  MoveL 1290 to (-200, -11.4, 56.6) mm, rotated rx 180 ry 0 rz 180 deg; joints [-15.315, -59.69, 128.134, 163.594, 69.246, -84.044]
  MoveL 1291 to (-200, -12, 56.6) mm, rotated rx 180 ry 0 rz 180 deg; joints [-15.315, -59.729, 128.133, 163.589, 69.207, -84.031]
  MoveL 1292 to (0, -12, 56.6) mm, rotated rx 180 ry 0 rz 180 deg; joints [-13.166, -51.617, 112.007, 164.94, 61.242, -82.624]
  MoveL 1293 to (0, -12.6, 56.6) mm, rotated rx 180 ry 0 rz 180 deg; joints [-13.166, -51.649, 112.006, 164.936, 61.21, -82.614]
  MoveL 1294 to (-200, -12.6, 56.6) mm, rotated rx 180 ry 0 rz 180 deg; joints [-15.315, -59.768, 128.131, 163.585, 69.169, -84.019]
  MoveL 1295 to (-200, -13.2, 56.6) mm, rotated rx 180 ry 0 rz 180 deg; joints [-15.315, -59.807, 128.13, 163.581, 69.13, -84.007]
  MoveL 1296 to (0, -13.2, 56.6) mm, rotated rx 180 ry 0 rz 180 deg; joints [-13.166, -51.681, 112.005, 164.931, 61.178, -82.605]
  MoveL 1297 to (0, -13.8, 56.6) mm, rotated rx 180 ry 0 rz 180 deg; joints [-13.166, -51.713, 112.003, 164.926, 61.146, -82.595]
  MoveL 1298 to (-200, -13.8, 56.6) mm, rotated rx 180 ry 0 rz 180 deg; joints [-15.315, -59.846, 128.129, 163.576, 69.091, -83.995]
  MoveL 1299 to (-200, -14.4, 56.6) mm, rotated rx 180 ry 0 rz 180 deg; joints [-15.315, -59.885, 128.127, 163.572, 69.052, -83.982]
  MoveL 1300 to (0, -14.4, 56.6) mm, rotated rx 180 ry 0 rz 180 deg; joints [-13.166, -51.745, 112.002, 164.921, 61.114, -82.585]
  MoveL 1301 to (0, -15, 56.6) mm, rotated rx 180 ry 0 rz 180 deg; joints [-13.166, -51.776, 112.001, 164.917, 61.082, -82.575]
  MoveL 1302 to (-200, -15, 56.6) mm, rotated rx 180 ry 0 rz 180 deg; joints [-15.315, -59.924, 128.126, 163.567, 69.013, -83.97]
  MoveL 1303 to (-200, -15.6, 56.6) mm, rotated rx 180 ry 0 rz 180 deg; joints [-15.315, -59.963, 128.124, 163.563, 68.975, -83.958]
  MoveL 1304 to (0, -15.6, 56.6) mm, rotated rx 180 ry 0 rz 180 deg; joints [-13.166, -51.808, 111.999, 164.912, 61.05, -82.565]
  MoveL 1305 to (0, -16.2, 56.6) mm, rotated rx 180 ry 0 rz 180 deg; joints [-13.166, -51.84, 111.998, 164.907, 61.018, -82.555]
  MoveL 1306 to (-200, -16.2, 56.6) mm, rotated rx 180 ry 0 rz 180 deg; joints [-15.315, -60.001, 128.122, 163.559, 68.936, -83.946]
  MoveL 1307 to (-200, -16.8, 56.6) mm, rotated rx 180 ry 0 rz 180 deg; joints [-15.315, -60.04, 128.121, 163.554, 68.897, -83.933]
  MoveL 1308 to (0, -16.8, 56.6) mm, rotated rx 180 ry 0 rz 180 deg; joints [-13.166, -51.872, 111.996, 164.902, 60.986, -82.545]
  MoveL 1309 to (0, -17.4, 56.6) mm, rotated rx 180 ry 0 rz 180 deg; joints [-13.166, -51.903, 111.995, 164.898, 60.954, -82.535]
  MoveL 1310 to (-200, -17.4, 56.6) mm, rotated rx 180 ry 0 rz 180 deg; joints [-15.315, -60.079, 128.119, 163.55, 68.858, -83.921]
  MoveL 1311 to (-200, -18, 56.6) mm, rotated rx 180 ry 0 rz 180 deg; joints [-15.315, -60.118, 128.117, 163.545, 68.819, -83.909]
  MoveL 1312 to (0, -18, 56.6) mm, rotated rx 180 ry 0 rz 180 deg; joints [-13.166, -51.935, 111.993, 164.893, 60.922, -82.526]
  MoveL 1313 to (0, -18.6, 56.6) mm, rotated rx 180 ry 0 rz 180 deg; joints [-13.166, -51.967, 111.992, 164.888, 60.89, -82.516]
  MoveL 1314 to (-200, -18.6, 56.6) mm, rotated rx 180 ry 0 rz 180 deg; joints [-15.315, -60.157, 128.116, 163.541, 68.78, -83.896]
  MoveL 1315 to (-200, -19.2, 56.6) mm, rotated rx 180 ry 0 rz 180 deg; joints [-15.315, -60.196, 128.114, 163.536, 68.741, -83.884]
  MoveL 1316 to (0, -19.2, 56.6) mm, rotated rx 180 ry 0 rz 180 deg; joints [-13.166, -51.998, 111.99, 164.883, 60.858, -82.506]
  MoveL 1317 to (0, -19.8, 56.6) mm, rotated rx 180 ry 0 rz 180 deg; joints [-13.166, -52.03, 111.988, 164.878, 60.826, -82.496]
  MoveL 1318 to (-200, -19.8, 56.6) mm, rotated rx 180 ry 0 rz 180 deg; joints [-15.315, -60.235, 128.112, 163.532, 68.702, -83.872]
  MoveL 1319 to (-200, -20.4, 56.6) mm, rotated rx 180 ry 0 rz 180 deg; joints [-15.315, -60.273, 128.11, 163.527, 68.663, -83.859]
  MoveL 1320 to (0, -20.4, 56.6) mm, rotated rx 180 ry 0 rz 180 deg; joints [-13.166, -52.062, 111.987, 164.873, 60.794, -82.486]
  MoveL 1321 to (0, -21, 56.6) mm, rotated rx 180 ry 0 rz 180 deg; joints [-13.166, -52.093, 111.985, 164.869, 60.762, -82.476]
  MoveL 1322 to (-200, -21, 56.6) mm, rotated rx 180 ry 0 rz 180 deg; joints [-15.315, -60.312, 128.108, 163.523, 68.624, -83.847]
  MoveL 1323 to (-200, -21.6, 56.6) mm, rotated rx 180 ry 0 rz 180 deg; joints [-15.315, -60.351, 128.107, 163.518, 68.585, -83.835]
  MoveL 1324 to (0, -21.6, 56.6) mm, rotated rx 180 ry 0 rz 180 deg; joints [-13.166, -52.125, 111.983, 164.864, 60.729, -82.466]
  MoveL 1325 to (0, -22.2, 56.6) mm, rotated rx 180 ry 0 rz 180 deg; joints [-13.166, -52.156, 111.982, 164.859, 60.697, -82.456]
  MoveL 1326 to (-200, -22.2, 56.6) mm, rotated rx 180 ry 0 rz 180 deg; joints [-15.315, -60.39, 128.105, 163.514, 68.546, -83.822]
  MoveL 1327 to (-200, -22.8, 56.6) mm, rotated rx 180 ry 0 rz 180 deg; joints [-15.315, -60.428, 128.103, 163.509, 68.507, -83.81]
  MoveL 1328 to (0, -22.8, 56.6) mm, rotated rx 180 ry 0 rz 180 deg; joints [-13.166, -52.188, 111.98, 164.854, 60.665, -82.446]
  MoveL 1329 to (0, -23.4, 56.6) mm, rotated rx 180 ry 0 rz 180 deg; joints [-13.166, -52.219, 111.978, 164.849, 60.633, -82.436]
  MoveL 1330 to (-200, -23.4, 56.6) mm, rotated rx 180 ry 0 rz 180 deg; joints [-15.315, -60.467, 128.101, 163.505, 68.468, -83.797]
  MoveL 1331 to (-200, -24, 56.6) mm, rotated rx 180 ry 0 rz 180 deg; joints [-15.315, -60.506, 128.099, 163.5, 68.429, -83.785]
  MoveL 1332 to (0, -24, 56.6) mm, rotated rx 180 ry 0 rz 180 deg; joints [-13.166, -52.251, 111.976, 164.844, 60.601, -82.426]
  MoveL 1333 to (0, -24.6, 56.6) mm, rotated rx 180 ry 0 rz 180 deg; joints [-13.166, -52.282, 111.974, 164.839, 60.568, -82.416]
  MoveL 1334 to (-200, -24.6, 56.6) mm, rotated rx 180 ry 0 rz 180 deg; joints [-15.315, -60.545, 128.097, 163.496, 68.39, -83.772]
  MoveL 1335 to (-200, -25.2, 56.6) mm, rotated rx 180 ry 0 rz 180 deg; joints [-15.315, -60.583, 128.095, 163.491, 68.351, -83.76]
  MoveL 1336 to (0, -25.2, 56.6) mm, rotated rx 180 ry 0 rz 180 deg; joints [-13.166, -52.314, 111.973, 164.834, 60.536, -82.406]
  MoveL 1337 to (0, -25.8, 56.6) mm, rotated rx 180 ry 0 rz 180 deg; joints [-13.166, -52.345, 111.971, 164.829, 60.504, -82.396]
  MoveL 1338 to (-200, -25.8, 56.6) mm, rotated rx 180 ry 0 rz 180 deg; joints [-15.315, -60.622, 128.092, 163.486, 68.312, -83.748]
  MoveL 1339 to (-200, -26.4, 56.6) mm, rotated rx 180 ry 0 rz 180 deg; joints [-15.315, -60.66, 128.09, 163.482, 68.273, -83.735]
  MoveL 1340 to (0, -26.4, 56.6) mm, rotated rx 180 ry 0 rz 180 deg; joints [-13.166, -52.377, 111.969, 164.824, 60.472, -82.386]
  MoveL 1341 to (0, -27, 56.6) mm, rotated rx 180 ry 0 rz 180 deg; joints [-13.166, -52.408, 111.967, 164.819, 60.439, -82.376]
  MoveL 1342 to (-200, -27, 56.6) mm, rotated rx 180 ry 0 rz 180 deg; joints [-15.315, -60.699, 128.088, 163.477, 68.234, -83.723]
  MoveL 1343 to (-200, -27.6, 56.6) mm, rotated rx 180 ry 0 rz 180 deg; joints [-15.315, -60.738, 128.086, 163.472, 68.195, -83.71]
  MoveL 1344 to (0, -27.6, 56.6) mm, rotated rx 180 ry 0 rz 180 deg; joints [-13.166, -52.44, 111.965, 164.814, 60.407, -82.366]
  MoveL 1345 to (0, -28.2, 56.6) mm, rotated rx 180 ry 0 rz 180 deg; joints [-13.166, -52.471, 111.963, 164.809, 60.375, -82.356]
  MoveL 1346 to (-200, -28.2, 56.6) mm, rotated rx 180 ry 0 rz 180 deg; joints [-15.315, -60.776, 128.084, 163.468, 68.156, -83.698]
  MoveL 1347 to (-200, -28.8, 56.6) mm, rotated rx 180 ry 0 rz 180 deg; joints [-15.315, -60.815, 128.081, 163.463, 68.116, -83.685]
  MoveL 1348 to (0, -28.8, 56.6) mm, rotated rx 180 ry 0 rz 180 deg; joints [-13.166, -52.503, 111.961, 164.804, 60.343, -82.346]
  MoveL 1349 to (0, -29.4, 56.6) mm, rotated rx 180 ry 0 rz 180 deg; joints [-13.166, -52.534, 111.959, 164.799, 60.31, -82.335]
  MoveL 1350 to (-200, -29.4, 56.6) mm, rotated rx 180 ry 0 rz 180 deg; joints [-15.315, -60.853, 128.079, 163.458, 68.077, -83.672]
  MoveL 1351 to (-200, -30, 56.6) mm, rotated rx 180 ry 0 rz 180 deg; joints [-15.315, -60.892, 128.077, 163.454, 68.038, -83.66]
  MoveL 1352 to (0, -30, 56.6) mm, rotated rx 180 ry 0 rz 180 deg; joints [-13.166, -52.565, 111.956, 164.794, 60.278, -82.325]
  MoveL 1353 to (0, -30.6, 56.58) mm, rotated rx 177.04 ry 0 rz 180 deg; joints [-13.235, -53.54, 111.838, 164.547, 59.233, -84.915]
  MoveL 1354 to (-200, -30.6, 56.58) mm, rotated rx 177.04 ry 0 rz 180 deg; joints [-15.394, -62.091, 127.948, 163.21, 66.774, -86.179]
  MoveL 1355 to (-200, -31.2, 56.54) mm, rotated rx 174.07 ry 0 rz 180 deg; joints [-15.428, -63.285, 127.806, 163.002, 65.501, -88.702]
  MoveL 1356 to (0, -31.2, 56.54) mm, rotated rx 174.07 ry 0 rz 180 deg; joints [-13.265, -54.511, 111.709, 164.333, 58.178, -87.515]
  MoveL 1357 to (0, -31.79, 56.46) mm, rotated rx 171.11 ry 0 rz 180 deg; joints [-13.255, -55.475, 111.57, 164.155, 57.114, -90.13]
  MoveL 1358 to (-200, -31.79, 56.46) mm, rotated rx 171.11 ry 0 rz 180 deg; joints [-15.417, -64.469, 127.651, 162.829, 64.219, -91.237]
  MoveL 1359 to (-200, -32.38, 56.35) mm, rotated rx 168.15 ry 0 rz 180 deg; joints [-15.36, -65.641, 127.484, 162.694, 62.932, -93.784]
  MoveL 1360 to (0, -32.38, 56.35) mm, rotated rx 168.15 ry 0 rz 180 deg; joints [-13.206, -56.43, 111.42, 164.013, 56.044, -92.762]
  MoveL 1361 to (0, -32.97, 56.21) mm, rotated rx 165.18 ry 0 rz 180 deg; joints [-13.118, -57.374, 111.26, 163.909, 54.969, -95.416]
  MoveL 1362 to (-200, -32.97, 56.21) mm, rotated rx 165.18 ry 0 rz 180 deg; joints [-15.259, -66.799, 127.305, 162.598, 61.643, -96.351]
  MoveL 1363 to (-200, -33.54, 56.05) mm, rotated rx 162.22 ry 0 rz 180 deg; joints [-15.112, -67.937, 127.115, 162.543, 60.354, -98.94]
  MoveL 1364 to (0, -33.54, 56.05) mm, rotated rx 162.22 ry 0 rz 180 deg; joints [-12.99, -58.304, 111.092, 163.846, 53.893, -98.094]
  MoveL 1365 to (0, -34.11, 55.85) mm, rotated rx 159.25 ry 0 rz 180 deg; joints [-12.824, -59.217, 110.914, 163.824, 52.818, -100.802]
  MoveL 1366 to (-200, -34.11, 55.85) mm, rotated rx 159.25 ry 0 rz 180 deg; joints [-14.921, -69.055, 126.916, 162.531, 59.067, -101.556]
  MoveL 1367 to (-200, -34.66, 55.62) mm, rotated rx 156.29 ry 0 rz 180 deg; joints [-14.686, -70.148, 126.706, 162.564, 57.786, -104.204]
  MoveL 1368 to (0, -34.66, 55.62) mm, rotated rx 156.29 ry 0 rz 180 deg; joints [-12.619, -60.112, 110.729, 163.847, 51.745, -103.542]
  MoveL 1369 to (0, -35.21, 55.37) mm, rotated rx 153.33 ry 0 rz 180 deg; joints [-12.376, -60.986, 110.538, 163.916, 50.677, -106.317]
  MoveL 1370 to (-200, -35.21, 55.37) mm, rotated rx 153.33 ry 0 rz 180 deg; joints [-14.406, -71.215, 126.489, 162.644, 56.513, -106.888]
  MoveL 1371 to (-200, -35.74, 55.08) mm, rotated rx 150.36 ry 0 rz 180 deg; joints [-14.083, -72.253, 126.264, 162.774, 55.251, -109.614]
  MoveL 1372 to (0, -35.74, 55.08) mm, rotated rx 150.36 ry 0 rz 180 deg; joints [-12.095, -61.837, 110.34, 164.034, 49.618, -109.135]
  MoveL 1373 to (0, -36.25, 54.77) mm, rotated rx 147.4 ry 0 rz 180 deg; joints [-11.777, -62.663, 110.136, 164.203, 48.57, -111.996]
  MoveL 1374 to (-200, -36.25, 54.77) mm, rotated rx 147.4 ry 0 rz 180 deg; joints [-13.716, -73.26, 126.033, 162.958, 54.004, -112.386]
  MoveL 1375 to (-200, -36.75, 54.44) mm, rotated rx 144.44 ry 0 rz 180 deg; joints [-13.307, -74.233, 125.797, 163.198, 52.775, -115.211]
  MoveL 1376 to (0, -36.75, 54.44) mm, rotated rx 144.44 ry 0 rz 180 deg; joints [-11.422, -63.463, 109.929, 164.427, 47.535, -114.907]
  MoveL 1377 to (0, -37.23, 54.08) mm, rotated rx 141.47 ry 0 rz 180 deg; joints [-11.032, -64.234, 109.719, 164.709, 46.517, -117.871]
  MoveL 1378 to (-200, -37.23, 54.08) mm, rotated rx 141.47 ry 0 rz 180 deg; joints [-12.856, -75.17, 125.557, 163.498, 51.566, -118.091]
  MoveL 1379 to (-200, -37.69, 53.69) mm, rotated rx 138.51 ry 0 rz 180 deg; joints [-12.364, -76.07, 125.315, 163.86, 50.381, -121.035]
  MoveL 1380 to (0, -37.69, 53.69) mm, rotated rx 138.51 ry 0 rz 180 deg; joints [-10.606, -64.975, 109.506, 165.05, 45.518, -120.893]
  MoveL 1381 to (0, -38.12, 53.28) mm, rotated rx 135.55 ry 0 rz 180 deg; joints [-10.146, -65.683, 109.292, 165.455, 44.542, -123.977]
  MoveL 1382 to (-200, -38.12, 53.28) mm, rotated rx 135.55 ry 0 rz 180 deg; joints [-11.832, -76.929, 125.071, 164.29, 49.223, -124.044]
  MoveL 1383 to (-200, -38.54, 52.85) mm, rotated rx 132.58 ry 0 rz 180 deg; joints [-11.261, -77.748, 124.828, 164.789, 48.098, -127.125]
  MoveL 1384 to (0, -38.54, 52.85) mm, rotated rx 132.58 ry 0 rz 180 deg; joints [-9.653, -66.359, 109.079, 165.925, 43.592, -127.125]
  MoveL 1385 to (0, -38.94, 52.4) mm, rotated rx 129.62 ry 0 rz 180 deg; joints [-9.128, -66.999, 108.867, 166.464, 42.671, -130.343]
  MoveL 1386 to (-200, -38.94, 52.4) mm, rotated rx 129.62 ry 0 rz 180 deg; joints [-10.652, -78.523, 124.586, 165.362, 47.007, -130.282]
  MoveL 1387 to (-200, -39.31, 51.92) mm, rotated rx 126.66 ry 0 rz 180 deg; joints [-10.007, -79.254, 124.348, 166.011, 45.956, -133.518]
  MoveL 1388 to (0, -39.31, 51.92) mm, rotated rx 126.66 ry 0 rz 180 deg; joints [-8.572, -67.603, 108.657, 167.074, 41.783, -133.633]
  MoveL 1389 to (0, -39.65, 51.44) mm, rotated rx 123.69 ry 0 rz 180 deg; joints [-7.986, -68.17, 108.45, 167.758, 40.932, -136.998]
  MoveL 1390 to (-200, -39.65, 51.44) mm, rotated rx 123.69 ry 0 rz 180 deg; joints [-9.326, -79.939, 124.113, 166.739, 44.949, -136.839]
  MoveL 1391 to (-200, -39.97, 50.93) mm, rotated rx 120.73 ry 0 rz 180 deg; joints [-8.612, -80.576, 123.885, 167.549, 43.99, -140.244]
  MoveL 1392 to (0, -39.97, 50.93) mm, rotated rx 120.73 ry 0 rz 180 deg; joints [-7.372, -68.697, 108.249, 168.515, 40.122, -140.44]
  MoveL 1393 to (0, -40.26, 50.4) mm, rotated rx 117.77 ry 0 rz 180 deg; joints [-6.731, -69.186, 108.053, 169.348, 39.355, -143.96]
  MoveL 1394 to (-200, -40.26, 50.4) mm, rotated rx 117.77 ry 0 rz 180 deg; joints [-7.867, -81.165, 123.663, 168.441, 43.084, -143.739]
  MoveL 1395 to (-200, -40.53, 49.87) mm, rotated rx 114.8 ry 0 rz 180 deg; joints [-7.091, -81.704, 123.45, 169.417, 42.234, -147.323]
  MoveL 1396 to (0, -40.53, 49.87) mm, rotated rx 114.8 ry 0 rz 180 deg; joints [-6.066, -69.633, 107.864, 170.256, 38.636, -147.559]
  MoveL 1397 to (0, -40.77, 49.31) mm, rotated rx 111.84 ry 0 rz 180 deg; joints [-5.378, -70.039, 107.683, 171.238, 37.97, -151.235]
  MoveL 1398 to (-200, -40.77, 49.31) mm, rotated rx 111.84 ry 0 rz 180 deg; joints [-6.288, -82.193, 123.246, 170.475, 41.447, -150.994]
  MoveL 1399 to (-200, -40.98, 48.75) mm, rotated rx 108.87 ry 0 rz 180 deg; joints [-5.46, -82.631, 123.053, 171.615, 40.726, -154.752]
  MoveL 1400 to (0, -40.98, 48.75) mm, rotated rx 108.87 ry 0 rz 180 deg; joints [-4.668, -70.402, 107.511, 172.293, 37.359, -154.987]
  MoveL 1401 to (0, -41.16, 48.18) mm, rotated rx 105.91 ry 0 rz 180 deg; joints [-3.939, -70.723, 107.349, 173.417, 36.808, -158.81]
  MoveL 1402 to (-200, -41.16, 48.18) mm, rotated rx 105.91 ry 0 rz 180 deg; joints [-4.608, -83.016, 122.871, 172.831, 40.077, -158.592]
  MoveL 1403 to (-200, -41.3, 47.6) mm, rotated rx 102.95 ry 0 rz 180 deg; joints [-3.736, -83.349, 122.703, 174.121, 39.502, -162.51]
  MoveL 1404 to (0, -41.3, 47.6) mm, rotated rx 102.95 ry 0 rz 180 deg; joints [-3.192, -71, 107.198, 174.605, 36.319, -162.701]
  MoveL 1405 to (0, -41.42, 47.01) mm, rotated rx 99.98 ry 0 rz 180 deg; joints [-2.431, -71.233, 107.058, 175.851, 35.897, -166.654]
  MoveL 1406 to (-200, -41.42, 47.01) mm, rotated rx 99.98 ry 0 rz 180 deg; joints [-2.845, -83.628, 122.548, 175.477, 39.007, -166.499]
  MoveL 1407 to (-200, -41.51, 46.42) mm, rotated rx 97.02 ry 0 rz 180 deg; joints [-1.94, -83.854, 122.408, 176.889, 38.595, -170.548]
  MoveL 1408 to (0, -41.51, 46.42) mm, rotated rx 97.02 ry 0 rz 180 deg; joints [-1.657, -71.421, 106.931, 177.148, 35.543, -170.659]
  MoveL 1409 to (0, -41.57, 45.82) mm, rotated rx 94.06 ry 0 rz 180 deg; joints [-0.873, -71.565, 106.816, 178.488, 35.261, -174.71]
  MoveL 1410 to (-200, -41.57, 45.82) mm, rotated rx 94.06 ry 0 rz 180 deg; joints [-1.022, -84.026, 122.283, 178.35, 38.268, -174.649]
  MoveL 1411 to (-200, -41.6, 45.22) mm, rotated rx 91.09 ry 0 rz 180 deg; joints [-0.094, -84.144, 122.173, 179.847, 38.029, -178.787]
  MoveL 1412 to (0, -41.6, 45.22) mm, rotated rx 91.09 ry 0 rz 180 deg; joints [-0.08, -71.664, 106.715, 179.86, 35.052, -178.793]
  MoveL 1413 to (0, -41.6, 44.62) mm, rotated rx 90 ry 0 rz 180 deg; joints [0.229, -71.689, 106.681, -179.6, 34.993, 179.672]
  MoveL 1414 to (-200, -41.6, 44.62) mm, rotated rx 90 ry 0 rz 180 deg; joints [0.268, -84.174, 122.137, -179.564, 37.964, 179.656]
  MoveL 1415 to (-200, -41.6, 44.02) mm, rotated rx 90 ry 0 rz 180 deg; joints [0.298, -84.174, 122.137, -179.516, 37.964, 179.618]
  MoveL 1416 to (0, -41.6, 44.02) mm, rotated rx 90 ry 0 rz 180 deg; joints [0.254, -71.689, 106.681, -179.556, 34.993, 179.637]
  MoveL 1417 to (0, -41.6, 43.42) mm, rotated rx 90 ry 0 rz 180 deg; joints [0.279, -71.688, 106.681, -179.513, 34.994, 179.601]
  MoveL 1418 to (-200, -41.6, 43.42) mm, rotated rx 90 ry 0 rz 180 deg; joints [0.327, -84.173, 122.137, -179.468, 37.965, 179.581]
  MoveL 1419 to (-200, -41.6, 42.82) mm, rotated rx 90 ry 0 rz 180 deg; joints [0.356, -84.173, 122.137, -179.42, 37.965, 179.543]
  MoveL 1420 to (0, -41.6, 42.82) mm, rotated rx 90 ry 0 rz 180 deg; joints [0.305, -71.688, 106.681, -179.469, 34.994, 179.565]
  MoveL 1421 to (0, -41.6, 42.22) mm, rotated rx 90 ry 0 rz 180 deg; joints [0.33, -71.688, 106.68, -179.425, 34.994, 179.529]
  MoveL 1422 to (-200, -41.6, 42.22) mm, rotated rx 90 ry 0 rz 180 deg; joints [0.386, -84.173, 122.136, -179.373, 37.965, 179.506]
  MoveL 1423 to (-200, -41.6, 41.62) mm, rotated rx 90 ry 0 rz 180 deg; joints [0.415, -84.173, 122.136, -179.325, 37.965, 179.468]
  MoveL 1424 to (0, -41.6, 41.62) mm, rotated rx 90 ry 0 rz 180 deg; joints [0.355, -71.688, 106.68, -179.382, 34.994, 179.493]
  MoveL 1425 to (0, -41.6, 41.02) mm, rotated rx 90 ry 0 rz 180 deg; joints [0.38, -71.687, 106.68, -179.338, 34.994, 179.458]
  MoveL 1426 to (-200, -41.6, 41.02) mm, rotated rx 90 ry 0 rz 180 deg; joints [0.444, -84.172, 122.136, -179.277, 37.965, 179.43]
  MoveL 1427 to (-200, -41.6, 40.42) mm, rotated rx 90 ry 0 rz 180 deg; joints [0.474, -84.172, 122.135, -179.23, 37.966, 179.393]
  MoveL 1428 to (0, -41.6, 40.42) mm, rotated rx 90 ry 0 rz 180 deg; joints [0.405, -71.687, 106.679, -179.294, 34.994, 179.422]
  MoveL 1429 to (0, -41.6, 39.82) mm, rotated rx 90 ry 0 rz 180 deg; joints [0.43, -71.687, 106.679, -179.251, 34.994, 179.386]
  MoveL 1430 to (-200, -41.6, 39.82) mm, rotated rx 90 ry 0 rz 180 deg; joints [0.503, -84.172, 122.135, -179.182, 37.966, 179.355]
  MoveL 1431 to (-200, -41.6, 39.22) mm, rotated rx 90 ry 0 rz 180 deg; joints [0.532, -84.171, 122.135, -179.134, 37.966, 179.318]
  MoveL 1432 to (0, -41.6, 39.22) mm, rotated rx 90 ry 0 rz 180 deg; joints [0.455, -71.687, 106.679, -179.207, 34.995, 179.35]
  MoveL 1433 to (0, -41.6, 38.62) mm, rotated rx 90 ry 0 rz 180 deg; joints [0.48, -71.686, 106.678, -179.163, 34.995, 179.314]
  MoveL 1434 to (-200, -41.6, 38.62) mm, rotated rx 90 ry 0 rz 180 deg; joints [0.562, -84.171, 122.134, -179.087, 37.967, 179.28]
  MoveL 1435 to (-200, -41.6, 38.02) mm, rotated rx 90 ry 0 rz 180 deg; joints [0.591, -84.171, 122.134, -179.039, 37.967, 179.242]
  MoveL 1436 to (0, -41.6, 38.02) mm, rotated rx 90 ry 0 rz 180 deg; joints [0.505, -71.686, 106.678, -179.119, 34.995, 179.279]
  MoveL 1437 to (0, -41.6, 37.42) mm, rotated rx 90 ry 0 rz 180 deg; joints [0.53, -71.686, 106.677, -179.076, 34.995, 179.243]
  MoveL 1438 to (-200, -41.6, 37.42) mm, rotated rx 90 ry 0 rz 180 deg; joints [0.62, -84.17, 122.133, -178.991, 37.967, 179.205]
  MoveL 1439 to (-200, -41.6, 36.82) mm, rotated rx 90 ry 0 rz 180 deg; joints [0.65, -84.17, 122.133, -178.944, 37.968, 179.167]
  MoveL 1440 to (0, -41.6, 36.82) mm, rotated rx 90 ry 0 rz 180 deg; joints [0.555, -71.685, 106.677, -179.032, 34.995, 179.207]
  MoveL 1441 to (0, -41.6, 36.22) mm, rotated rx 90 ry 0 rz 180 deg; joints [0.58, -71.685, 106.676, -178.988, 34.996, 179.171]
  MoveL 1442 to (-200, -41.6, 36.22) mm, rotated rx 90 ry 0 rz 180 deg; joints [0.679, -84.169, 122.132, -178.896, 37.968, 179.13]
  MoveL 1443 to (-200, -41.6, 35.62) mm, rotated rx 90 ry 0 rz 180 deg; joints [0.708, -84.169, 122.132, -178.848, 37.968, 179.092]
  MoveL 1444 to (0, -41.6, 35.62) mm, rotated rx 90 ry 0 rz 180 deg; joints [0.605, -71.685, 106.676, -178.945, 34.996, 179.135]
  MoveL 1445 to (0, -41.6, 35.02) mm, rotated rx 90 ry 0 rz 180 deg; joints [0.63, -71.684, 106.675, -178.901, 34.996, 179.1]
  MoveL 1446 to (-200, -41.6, 35.02) mm, rotated rx 90 ry 0 rz 180 deg; joints [0.738, -84.168, 122.131, -178.801, 37.969, 179.055]
  MoveL 1447 to (-200, -41.6, 34.42) mm, rotated rx 90 ry 0 rz 180 deg; joints [0.767, -84.168, 122.131, -178.753, 37.969, 179.017]
  MoveL 1448 to (0, -41.6, 34.42) mm, rotated rx 90 ry 0 rz 180 deg; joints [0.655, -71.684, 106.675, -178.857, 34.996, 179.064]
  MoveL 1449 to (0, -41.6, 33.82) mm, rotated rx 90 ry 0 rz 180 deg; joints [0.68, -71.683, 106.674, -178.814, 34.997, 179.028]
  MoveL 1450 to (-200, -41.6, 33.82) mm, rotated rx 90 ry 0 rz 180 deg; joints [0.796, -84.167, 122.13, -178.705, 37.97, 178.979]
  MoveL 1451 to (-200, -41.6, 33.22) mm, rotated rx 90 ry 0 rz 180 deg; joints [0.826, -84.167, 122.129, -178.658, 37.97, 178.942]
  MoveL 1452 to (0, -41.6, 33.22) mm, rotated rx 90 ry 0 rz 180 deg; joints [0.705, -71.683, 106.674, -178.77, 34.997, 178.992]
  MoveL 1453 to (0, -41.6, 32.62) mm, rotated rx 90 ry 0 rz 180 deg; joints [0.73, -71.682, 106.673, -178.726, 34.997, 178.957]
  MoveL 1454 to (-200, -41.6, 32.62) mm, rotated rx 90 ry 0 rz 180 deg; joints [0.855, -84.166, 122.129, -178.61, 37.971, 178.904]
  MoveL 1455 to (-200, -41.6, 32.02) mm, rotated rx 90 ry 0 rz 180 deg; joints [0.884, -84.166, 122.128, -178.562, 37.971, 178.867]
  MoveL 1456 to (0, -41.6, 32.02) mm, rotated rx 90 ry 0 rz 180 deg; joints [0.756, -71.682, 106.672, -178.683, 34.997, 178.921]
  MoveL 1457 to (0, -41.6, 31.42) mm, rotated rx 90 ry 0 rz 180 deg; joints [0.781, -71.682, 106.672, -178.639, 34.998, 178.885]
  MoveL 1458 to (-200, -41.6, 31.42) mm, rotated rx 90 ry 0 rz 180 deg; joints [0.914, -84.165, 122.127, -178.515, 37.972, 178.829]
  MoveL 1459 to (-200, -41.6, 30.82) mm, rotated rx 90 ry 0 rz 180 deg; joints [0.943, -84.164, 122.127, -178.467, 37.972, 178.792]
  MoveL 1460 to (0, -41.6, 30.82) mm, rotated rx 90 ry 0 rz 180 deg; joints [0.806, -71.681, 106.671, -178.595, 34.998, 178.849]
  MoveL 1461 to (0, -41.6, 30.22) mm, rotated rx 90 ry 0 rz 180 deg; joints [0.831, -71.68, 106.67, -178.552, 34.998, 178.813]
  MoveL 1462 to (-200, -41.6, 30.22) mm, rotated rx 90 ry 0 rz 180 deg; joints [0.972, -84.164, 122.126, -178.419, 37.973, 178.754]
  MoveL 1463 to (-200, -41.6, 29.62) mm, rotated rx 90 ry 0 rz 180 deg; joints [1.002, -84.163, 122.125, -178.372, 37.973, 178.716]
  MoveL 1464 to (0, -41.6, 29.62) mm, rotated rx 90 ry 0 rz 180 deg; joints [0.856, -71.68, 106.67, -178.508, 34.999, 178.778]
  MoveL 1465 to (0, -41.6, 29.02) mm, rotated rx 90 ry 0 rz 180 deg; joints [0.881, -71.679, 106.669, -178.464, 34.999, 178.742]
  MoveL 1466 to (-200, -41.6, 29.02) mm, rotated rx 90 ry 0 rz 180 deg; joints [1.031, -84.163, 122.125, -178.324, 37.974, 178.679]
  MoveL 1467 to (-200, -41.6, 28.42) mm, rotated rx 90 ry 0 rz 180 deg; joints [1.06, -84.162, 122.124, -178.277, 37.975, 178.641]
  MoveL 1468 to (0, -41.6, 28.42) mm, rotated rx 90 ry 0 rz 180 deg; joints [0.906, -71.679, 106.668, -178.421, 34.999, 178.706]
  MoveL 1469 to (0, -41.6, 27.82) mm, rotated rx 90 ry 0 rz 180 deg; joints [0.931, -71.678, 106.667, -178.377, 35, 178.67]
  MoveL 1470 to (-200, -41.6, 27.82) mm, rotated rx 90 ry 0 rz 180 deg; joints [1.09, -84.161, 122.123, -178.229, 37.975, 178.604]
  MoveL 1471 to (-200, -41.6, 27.22) mm, rotated rx 90 ry 0 rz 180 deg; joints [1.119, -84.16, 122.122, -178.181, 37.976, 178.566]
  MoveL 1472 to (0, -41.6, 27.22) mm, rotated rx 90 ry 0 rz 180 deg; joints [0.956, -71.678, 106.666, -178.333, 35, 178.635]
  MoveL 1473 to (0, -41.6, 26.62) mm, rotated rx 90 ry 0 rz 180 deg; joints [0.981, -71.677, 106.666, -178.29, 35.001, 178.599]
  MoveL 1474 to (-200, -41.6, 26.62) mm, rotated rx 90 ry 0 rz 180 deg; joints [1.148, -84.16, 122.121, -178.134, 37.976, 178.529]
  MoveL 1475 to (-200, -41.6, 26.02) mm, rotated rx 90 ry 0 rz 180 deg; joints [1.178, -84.159, 122.12, -178.086, 37.977, 178.491]
  MoveL 1476 to (0, -41.6, 26.02) mm, rotated rx 90 ry 0 rz 180 deg; joints [1.006, -71.676, 106.665, -178.246, 35.001, 178.563]
  MoveL 1477 to (0, -41.6, 25.42) mm, rotated rx 90 ry 0 rz 180 deg; joints [1.031, -71.676, 106.664, -178.202, 35.001, 178.527]
  MoveL 1478 to (-200, -41.6, 25.42) mm, rotated rx 90 ry 0 rz 180 deg; joints [1.207, -84.158, 122.119, -178.038, 37.978, 178.453]
  MoveL 1479 to (-200, -41.6, 24.82) mm, rotated rx 90 ry 0 rz 180 deg; joints [1.236, -84.157, 122.119, -177.991, 37.978, 178.416]
  MoveL 1480 to (0, -41.6, 24.82) mm, rotated rx 90 ry 0 rz 180 deg; joints [1.056, -71.675, 106.663, -178.159, 35.002, 178.491]
  MoveL 1481 to (0, -41.6, 24.22) mm, rotated rx 90 ry 0 rz 180 deg; joints [1.081, -71.674, 106.662, -178.115, 35.002, 178.456]
  MoveL 1482 to (-200, -41.6, 24.22) mm, rotated rx 90 ry 0 rz 180 deg; joints [1.266, -84.156, 122.118, -177.943, 37.979, 178.378]
  MoveL 1483 to (-200, -41.6, 23.62) mm, rotated rx 90 ry 0 rz 180 deg; joints [1.295, -84.155, 122.117, -177.895, 37.98, 178.341]
  MoveL 1484 to (0, -41.6, 23.62) mm, rotated rx 90 ry 0 rz 180 deg; joints [1.106, -71.674, 106.661, -178.071, 35.003, 178.42]
  MoveL 1485 to (0, -41.6, 23.02) mm, rotated rx 90 ry 0 rz 180 deg; joints [1.131, -71.673, 106.66, -178.028, 35.003, 178.384]
  MoveL 1486 to (-200, -41.6, 23.02) mm, rotated rx 90 ry 0 rz 180 deg; joints [1.324, -84.155, 122.116, -177.848, 37.981, 178.303]
  MoveL 1487 to (-200, -41.6, 22.42) mm, rotated rx 90 ry 0 rz 180 deg; joints [1.354, -84.154, 122.115, -177.8, 37.981, 178.266]
  MoveL 1488 to (0, -41.6, 22.42) mm, rotated rx 90 ry 0 rz 180 deg; joints [1.156, -71.672, 106.659, -177.984, 35.004, 178.348]
  MoveL 1489 to (0, -41.6, 21.82) mm, rotated rx 90 ry 0 rz 180 deg; joints [1.181, -71.671, 106.658, -177.94, 35.004, 178.313]
  MoveL 1490 to (-200, -41.6, 21.82) mm, rotated rx 90 ry 0 rz 180 deg; joints [1.383, -84.153, 122.114, -177.753, 37.982, 178.228]
  MoveL 1491 to (-200, -41.6, 21.22) mm, rotated rx 90 ry 0 rz 180 deg; joints [1.412, -84.152, 122.113, -177.705, 37.983, 178.191]
  MoveL 1492 to (0, -41.6, 21.22) mm, rotated rx 90 ry 0 rz 180 deg; joints [1.206, -71.671, 106.657, -177.897, 35.004, 178.277]
  MoveL 1493 to (0, -41.6, 20.62) mm, rotated rx 90 ry 0 rz 180 deg; joints [1.231, -71.67, 106.656, -177.853, 35.005, 178.241]
  MoveL 1494 to (-200, -41.6, 20.62) mm, rotated rx 90 ry 0 rz 180 deg; joints [1.442, -84.151, 122.111, -177.657, 37.984, 178.153]
  MoveL 1495 to (-200, -41.6, 20.02) mm, rotated rx 90 ry 0 rz 180 deg; joints [1.471, -84.15, 122.11, -177.61, 37.985, 178.116]
  MoveL 1496 to (0, -41.6, 20.02) mm, rotated rx 90 ry 0 rz 180 deg; joints [1.257, -71.669, 106.655, -177.809, 35.005, 178.205]
  MoveL 1497 to (0, -41.6, 19.42) mm, rotated rx 90 ry 0 rz 180 deg; joints [1.282, -71.668, 106.654, -177.766, 35.006, 178.17]
  MoveL 1498 to (-200, -41.6, 19.42) mm, rotated rx 90 ry 0 rz 180 deg; joints [1.5, -84.149, 122.109, -177.562, 37.986, 178.078]
  MoveL 1499 to (-200, -41.6, 18.82) mm, rotated rx 90 ry 0 rz 180 deg; joints [1.529, -84.148, 122.108, -177.514, 37.986, 178.041]
  MoveL 1500 to (0, -41.6, 18.82) mm, rotated rx 90 ry 0 rz 180 deg; joints [1.307, -71.667, 106.653, -177.722, 35.006, 178.134]
  MoveL 1501 to (0, -41.6, 18.22) mm, rotated rx 90 ry 0 rz 180 deg; joints [1.332, -71.667, 106.651, -177.678, 35.007, 178.098]
  MoveL 1502 to (-200, -41.6, 18.22) mm, rotated rx 90 ry 0 rz 180 deg; joints [1.559, -84.147, 122.107, -177.467, 37.987, 178.003]
  MoveL 1503 to (-200, -41.6, 17.62) mm, rotated rx 90 ry 0 rz 180 deg; joints [1.588, -84.146, 122.106, -177.419, 37.988, 177.966]
  MoveL 1504 to (0, -41.6, 17.62) mm, rotated rx 90 ry 0 rz 180 deg; joints [1.357, -71.666, 106.65, -177.635, 35.008, 178.062]
  MoveL 1505 to (0, -41.6, 17.02) mm, rotated rx 90 ry 0 rz 180 deg; joints [1.382, -71.665, 106.649, -177.591, 35.008, 178.027]
  MoveL 1506 to (-200, -41.6, 17.02) mm, rotated rx 90 ry 0 rz 180 deg; joints [1.617, -84.145, 122.105, -177.372, 37.989, 177.928]
  MoveL 1507 to (-200, -41.6, 16.42) mm, rotated rx 90 ry 0 rz 180 deg; joints [1.647, -84.144, 122.103, -177.324, 37.99, 177.891]
  MoveL 1508 to (0, -41.6, 16.42) mm, rotated rx 90 ry 0 rz 180 deg; joints [1.407, -71.664, 106.648, -177.547, 35.009, 177.991]
  MoveL 1509 to (0, -41.6, 15.82) mm, rotated rx 90 ry 0 rz 180 deg; joints [1.432, -71.663, 106.647, -177.504, 35.009, 177.955]
  MoveL 1510 to (-200, -41.6, 15.82) mm, rotated rx 90 ry 0 rz 180 deg; joints [1.676, -84.142, 122.102, -177.277, 37.991, 177.853]
  MoveL 1511 to (-200, -41.6, 15.22) mm, rotated rx 90 ry 0 rz 180 deg; joints [1.705, -84.141, 122.101, -177.229, 37.992, 177.815]
  MoveL 1512 to (0, -41.6, 15.22) mm, rotated rx 90 ry 0 rz 180 deg; joints [1.457, -71.662, 106.645, -177.46, 35.01, 177.919]
  MoveL 1513 to (0, -41.59, 14.62) mm, rotated rx 88.13 ry 0 rz 180 deg; joints [1.97, -71.674, 106.57, -176.559, 34.944, 175.307]
  MoveL 1514 to (-200, -41.59, 14.62) mm, rotated rx 88.13 ry 0 rz 180 deg; joints [2.306, -84.155, 122.022, -176.247, 37.926, 175.167]
  MoveL 1515 to (-200, -41.56, 14.02) mm, rotated rx 85.17 ry 0 rz 180 deg; joints [3.242, -84.133, 121.91, -174.717, 37.896, 170.993]
  MoveL 1516 to (0, -41.56, 14.02) mm, rotated rx 85.17 ry 0 rz 180 deg; joints [2.77, -71.657, 106.462, -175.155, 34.901, 171.189]
  MoveL 1517 to (0, -41.49, 13.43) mm, rotated rx 82.2 ry 0 rz 180 deg; joints [3.571, -71.595, 106.369, -173.756, 34.934, 167.076]
  MoveL 1518 to (-200, -41.49, 13.43) mm, rotated rx 82.2 ry 0 rz 180 deg; joints [4.178, -84.057, 121.816, -173.197, 37.955, 166.828]
  MoveL 1519 to (-200, -41.4, 12.83) mm, rotated rx 79.24 ry 0 rz 180 deg; joints [5.111, -83.928, 121.739, -171.699, 38.104, 162.689]
  MoveL 1520 to (0, -41.4, 12.83) mm, rotated rx 79.24 ry 0 rz 180 deg; joints [4.369, -71.488, 106.29, -172.375, 35.041, 162.983]
  MoveL 1521 to (0, -41.27, 12.25) mm, rotated rx 76.28 ry 0 rz 180 deg; joints [5.163, -71.337, 106.227, -171.024, 35.221, 158.922]
  MoveL 1522 to (-200, -41.27, 12.25) mm, rotated rx 76.28 ry 0 rz 180 deg; joints [6.038, -83.745, 121.679, -170.238, 38.34, 158.589]
  MoveL 1523 to (-200, -41.11, 11.67) mm, rotated rx 73.31 ry 0 rz 180 deg; joints [6.956, -83.51, 121.636, -168.822, 38.66, 154.54]
  MoveL 1524 to (0, -41.11, 11.67) mm, rotated rx 73.31 ry 0 rz 180 deg; joints [5.949, -71.142, 106.178, -169.711, 35.473, 154.902]
  MoveL 1525 to (0, -40.92, 11.1) mm, rotated rx 70.35 ry 0 rz 180 deg; joints [6.727, -70.905, 106.144, -168.447, 35.794, 150.934]
  MoveL 1526 to (-200, -40.92, 11.1) mm, rotated rx 70.35 ry 0 rz 180 deg; joints [7.861, -83.224, 121.611, -167.464, 39.062, 150.553]
  MoveL 1527 to (-200, -40.71, 10.54) mm, rotated rx 67.38 ry 0 rz 180 deg; joints [8.753, -82.886, 121.602, -166.171, 39.541, 146.635]
  MoveL 1528 to (0, -40.71, 10.54) mm, rotated rx 67.38 ry 0 rz 180 deg; joints [7.492, -70.624, 106.125, -167.239, 36.181, 147.025]
  MoveL 1529 to (0, -40.46, 9.99) mm, rotated rx 64.42 ry 0 rz 180 deg; joints [8.244, -70.302, 106.12, -166.094, 36.63, 143.184]
  MoveL 1530 to (-200, -40.46, 9.99) mm, rotated rx 64.42 ry 0 rz 180 deg; joints [9.626, -82.499, 121.609, -164.951, 40.093, 142.798]
  MoveL 1531 to (-200, -40.19, 9.46) mm, rotated rx 61.46 ry 0 rz 180 deg; joints [10.481, -82.062, 121.633, -163.807, 40.714, 139.043]
  MoveL 1532 to (0, -40.19, 9.46) mm, rotated rx 61.46 ry 0 rz 180 deg; joints [8.98, -69.938, 106.129, -165.017, 37.139, 139.414]
  MoveL 1533 to (0, -39.89, 8.94) mm, rotated rx 58.49 ry 0 rz 180 deg; joints [9.698, -69.535, 106.151, -164.012, 37.704, 135.721]
  MoveL 1534 to (-200, -39.89, 8.94) mm, rotated rx 58.49 ry 0 rz 180 deg; joints [11.313, -81.577, 121.671, -162.744, 41.399, 135.376]
  MoveL 1535 to (-200, -39.56, 8.44) mm, rotated rx 55.53 ry 0 rz 180 deg; joints [12.121, -81.046, 121.724, -161.764, 42.143, 131.801]
  MoveL 1536 to (0, -39.56, 8.44) mm, rotated rx 55.53 ry 0 rz 180 deg; joints [10.396, -69.092, 106.187, -163.082, 38.321, 132.108]
  MoveL 1537 to (0, -39.21, 7.95) mm, rotated rx 52.57 ry 0 rz 180 deg; joints [11.072, -68.611, 106.235, -162.227, 38.986, 128.575]
  MoveL 1538 to (-200, -39.21, 7.95) mm, rotated rx 52.57 ry 0 rz 180 deg; joints [12.902, -80.469, 121.791, -160.867, 42.942, 128.316]
  MoveL 1539 to (-200, -38.83, 7.48) mm, rotated rx 49.6 ry 0 rz 180 deg; joints [13.655, -79.847, 121.871, -160.054, 43.791, 124.923]
  MoveL 1540 to (0, -38.83, 7.48) mm, rotated rx 49.6 ry 0 rz 180 deg; joints [11.724, -68.093, 106.295, -161.449, 39.696, 125.125]
  MoveL 1541 to (0, -38.43, 7.04) mm, rotated rx 46.64 ry 0 rz 180 deg; joints [12.352, -67.539, 106.366, -160.747, 40.446, 121.754]
  MoveL 1542 to (-200, -38.43, 7.04) mm, rotated rx 46.64 ry 0 rz 180 deg; joints [14.378, -79.182, 121.964, -159.322, 44.687, 121.618]
  MoveL 1543 to (-200, -38.01, 6.61) mm, rotated rx 43.68 ry 0 rz 180 deg; joints [15.07, -78.476, 122.067, -158.669, 45.623, 118.401]
  MoveL 1544 to (0, -38.01, 6.61) mm, rotated rx 43.68 ry 0 rz 180 deg; joints [12.953, -66.951, 106.447, -160.119, 41.233, 118.462]
  MoveL 1545 to (0, -37.57, 6.21) mm, rotated rx 40.71 ry 0 rz 180 deg; joints [13.526, -66.329, 106.538, -159.563, 42.054, 115.246]
  MoveL 1546 to (-200, -37.57, 6.21) mm, rotated rx 40.71 ry 0 rz 180 deg; joints [15.728, -77.73, 122.181, -158.093, 46.597, 115.266]
  MoveL 1547 to (-200, -37.1, 5.83) mm, rotated rx 37.75 ry 0 rz 180 deg; joints [16.351, -76.945, 122.304, -157.591, 47.605, 112.211]
  MoveL 1548 to (0, -37.1, 5.83) mm, rotated rx 37.75 ry 0 rz 180 deg; joints [14.07, -65.675, 106.638, -159.078, 42.906, 112.104]
  MoveL 1549 to (0, -36.62, 5.47) mm, rotated rx 34.78 ry 0 rz 180 deg; joints [14.583, -64.99, 106.746, -158.661, 43.783, 109.034]
  MoveL 1550 to (-200, -36.62, 5.47) mm, rotated rx 34.78 ry 0 rz 180 deg; joints [16.939, -76.123, 122.435, -157.16, 48.642, 109.233]
  MoveL 1551 to (-200, -36.12, 5.14) mm, rotated rx 31.82 ry 0 rz 180 deg; joints [17.49, -75.265, 122.574, -156.794, 49.706, 106.325]
  MoveL 1552 to (0, -36.12, 5.14) mm, rotated rx 31.82 ry 0 rz 180 deg; joints [15.066, -64.276, 106.861, -158.308, 44.686, 106.029]
  MoveL 1553 to (0, -35.6, 4.84) mm, rotated rx 28.86 ry 0 rz 180 deg; joints [15.515, -63.535, 106.982, -158.016, 45.608, 103.088]
  MoveL 1554 to (-200, -35.6, 4.84) mm, rotated rx 28.86 ry 0 rz 180 deg; joints [18.004, -74.375, 122.719, -156.492, 50.794, 103.484]
  MoveL 1555 to (-200, -35.07, 4.57) mm, rotated rx 25.89 ry 0 rz 180 deg; joints [18.478, -73.452, 122.869, -156.25, 51.902, 100.705]
  MoveL 1556 to (0, -35.07, 4.57) mm, rotated rx 25.89 ry 0 rz 180 deg; joints [15.932, -62.768, 107.108, -157.784, 46.55, 100.205]
  MoveL 1557 to (0, -34.52, 4.32) mm, rotated rx 22.93 ry 0 rz 180 deg; joints [16.315, -61.976, 107.24, -157.606, 47.507, 97.377]
  MoveL 1558 to (-200, -34.52, 4.32) mm, rotated rx 22.93 ry 0 rz 180 deg; joints [18.914, -72.5, 123.023, -156.063, 53.027, 97.982]
  MoveL 1559 to (-200, -33.96, 4.1) mm, rotated rx 19.97 ry 0 rz 180 deg; joints [19.309, -71.52, 123.181, -155.929, 54.167, 95.312]
  MoveL 1560 to (0, -33.96, 4.1) mm, rotated rx 19.97 ry 0 rz 180 deg; joints [16.663, -61.161, 107.374, -157.481, 48.477, 94.599]
  MoveL 1561 to (0, -33.39, 3.91) mm, rotated rx 17 ry 0 rz 180 deg; joints [16.975, -60.326, 107.512, -157.406, 49.458, 91.868]
  MoveL 1562 to (-200, -33.39, 3.91) mm, rotated rx 17 ry 0 rz 180 deg; joints [19.665, -70.514, 123.341, -155.845, 55.32, 92.688]
  MoveL 1563 to (-200, -32.81, 3.75) mm, rotated rx 14.04 ry 0 rz 180 deg; joints [19.979, -69.484, 123.502, -155.807, 56.484, 90.107]
  MoveL 1564 to (0, -32.81, 3.75) mm, rotated rx 14.04 ry 0 rz 180 deg; joints [17.252, -59.471, 107.652, -157.378, 50.448, 89.179]
  MoveL 1565 to (0, -32.23, 3.62) mm, rotated rx 11.08 ry 0 rz 180 deg; joints [17.493, -58.599, 107.794, -157.394, 51.445, 86.528]
  MoveL 1566 to (-200, -32.23, 3.62) mm, rotated rx 11.08 ry 0 rz 180 deg; joints [20.252, -68.433, 123.664, -155.813, 57.655, 87.564]
  MoveL 1567 to (-200, -31.64, 3.52) mm, rotated rx 8.11 ry 0 rz 180 deg; joints [20.483, -67.362, 123.825, -155.86, 58.832, 85.055]
  MoveL 1568 to (0, -31.64, 3.52) mm, rotated rx 8.11 ry 0 rz 180 deg; joints [17.698, -57.712, 107.936, -157.452, 52.446, 83.912]
  MoveL 1569 to (0, -31.04, 3.45) mm, rotated rx 5.15 ry 0 rz 180 deg; joints [17.865, -56.811, 108.078, -157.55, 53.45, 81.325]
  MoveL 1570 to (-200, -31.04, 3.45) mm, rotated rx 5.15 ry 0 rz 180 deg; joints [20.673, -66.274, 123.986, -155.946, 60.014, 82.573]
  MoveL 1571 to (-200, -30.44, 3.41) mm, rotated rx 2.19 ry 0 rz 180 deg; joints [20.821, -65.172, 124.144, -156.07, 61.198, 80.118]
  MoveL 1572 to (0, -30.44, 3.41) mm, rotated rx 2.19 ry 0 rz 180 deg; joints [17.996, -55.9, 108.22, -157.685, 54.455, 78.766]
  MoveL 1573 to (0, -29.84, 3.4) mm, rotated rx 0 ry 0 rz 180 deg; joints [18.068, -55.214, 108.325, -157.81, 55.204, 76.897]
  MoveL 1574 to (-200, -29.84, 3.4) mm, rotated rx 0 ry 0 rz 180 deg; joints [20.902, -64.342, 124.261, -156.186, 62.081, 78.324]
  MoveL 1575 to (-200, -29.24, 3.4) mm, rotated rx 0 ry 0 rz 180 deg; joints [20.902, -64.308, 124.268, -156.195, 62.118, 78.343]
  MoveL 1576 to (0, -29.24, 3.4) mm, rotated rx 0 ry 0 rz 180 deg; joints [18.068, -55.186, 108.332, -157.819, 55.235, 76.912]
  MoveL 1577 to (0, -28.64, 3.4) mm, rotated rx 0 ry 0 rz 180 deg; joints [18.068, -55.158, 108.338, -157.828, 55.267, 76.928]
  MoveL 1578 to (-200, -28.64, 3.4) mm, rotated rx 0 ry 0 rz 180 deg; joints [20.902, -64.274, 124.275, -156.203, 62.155, 78.361]
  MoveL 1579 to (-200, -28.04, 3.4) mm, rotated rx 0 ry 0 rz 180 deg; joints [20.902, -64.24, 124.282, -156.212, 62.193, 78.38]
  MoveL 1580 to (0, -28.04, 3.4) mm, rotated rx 0 ry 0 rz 180 deg; joints [18.068, -55.13, 108.344, -157.837, 55.299, 76.944]
  MoveL 1581 to (0, -27.44, 3.4) mm, rotated rx 0 ry 0 rz 180 deg; joints [18.068, -55.102, 108.35, -157.846, 55.331, 76.96]
  MoveL 1582 to (-200, -27.44, 3.4) mm, rotated rx 0 ry 0 rz 180 deg; joints [20.902, -64.206, 124.289, -156.221, 62.23, 78.399]
  MoveL 1583 to (-200, -26.84, 3.4) mm, rotated rx 0 ry 0 rz 180 deg; joints [20.902, -64.172, 124.295, -156.229, 62.267, 78.417]
  MoveL 1584 to (0, -26.84, 3.4) mm, rotated rx 0 ry 0 rz 180 deg; joints [18.068, -55.074, 108.357, -157.854, 55.362, 76.975]
  MoveL 1585 to (0, -26.24, 3.4) mm, rotated rx 0 ry 0 rz 180 deg; joints [18.068, -55.046, 108.363, -157.863, 55.394, 76.991]
  MoveL 1586 to (-200, -26.24, 3.4) mm, rotated rx 0 ry 0 rz 180 deg; joints [20.902, -64.138, 124.302, -156.238, 62.305, 78.436]
  MoveL 1587 to (-200, -25.64, 3.4) mm, rotated rx 0 ry 0 rz 180 deg; joints [20.902, -64.104, 124.309, -156.246, 62.342, 78.454]
  MoveL 1588 to (0, -25.64, 3.4) mm, rotated rx 0 ry 0 rz 180 deg; joints [18.068, -55.018, 108.369, -157.872, 55.426, 77.007]
  MoveL 1589 to (0, -25.04, 3.4) mm, rotated rx 0 ry 0 rz 180 deg; joints [18.068, -54.99, 108.375, -157.881, 55.457, 77.022]
  MoveL 1590 to (-200, -25.04, 3.4) mm, rotated rx 0 ry 0 rz 180 deg; joints [20.902, -64.069, 124.315, -156.255, 62.379, 78.473]
  MoveL 1591 to (-200, -24.44, 3.4) mm, rotated rx 0 ry 0 rz 180 deg; joints [20.902, -64.035, 124.322, -156.264, 62.417, 78.491]
  MoveL 1592 to (0, -24.44, 3.4) mm, rotated rx 0 ry 0 rz 180 deg; joints [18.068, -54.962, 108.381, -157.89, 55.489, 77.038]
  MoveL 1593 to (0, -23.84, 3.4) mm, rotated rx 0 ry 0 rz 180 deg; joints [18.068, -54.934, 108.387, -157.899, 55.521, 77.053]
  MoveL 1594 to (-200, -23.84, 3.4) mm, rotated rx 0 ry 0 rz 180 deg; joints [20.902, -64.001, 124.329, -156.272, 62.454, 78.51]
  MoveL 1595 to (-200, -23.24, 3.4) mm, rotated rx 0 ry 0 rz 180 deg; joints [20.902, -63.967, 124.335, -156.281, 62.491, 78.528]
  MoveL 1596 to (0, -23.24, 3.4) mm, rotated rx 0 ry 0 rz 180 deg; joints [18.068, -54.906, 108.393, -157.908, 55.552, 77.069]
  MoveL 1597 to (0, -22.64, 3.4) mm, rotated rx 0 ry 0 rz 180 deg; joints [18.068, -54.877, 108.399, -157.916, 55.584, 77.085]
  MoveL 1598 to (-200, -22.64, 3.4) mm, rotated rx 0 ry 0 rz 180 deg; joints [20.902, -63.933, 124.342, -156.289, 62.528, 78.547]
  MoveL 1599 to (-200, -22.04, 3.4) mm, rotated rx 0 ry 0 rz 180 deg; joints [20.902, -63.899, 124.348, -156.298, 62.566, 78.565]
  MoveL 1600 to (0, -22.04, 3.4) mm, rotated rx 0 ry 0 rz 180 deg; joints [18.068, -54.849, 108.405, -157.925, 55.615, 77.1]
  MoveL 1601 to (0, -21.44, 3.4) mm, rotated rx 0 ry 0 rz 180 deg; joints [18.068, -54.821, 108.411, -157.934, 55.647, 77.116]
  MoveL 1602 to (-200, -21.44, 3.4) mm, rotated rx 0 ry 0 rz 180 deg; joints [20.902, -63.864, 124.355, -156.306, 62.603, 78.584]
  MoveL 1603 to (-200, -20.84, 3.4) mm, rotated rx 0 ry 0 rz 180 deg; joints [20.902, -63.83, 124.361, -156.315, 62.64, 78.602]
  MoveL 1604 to (0, -20.84, 3.4) mm, rotated rx 0 ry 0 rz 180 deg; joints [18.068, -54.793, 108.417, -157.943, 55.679, 77.131]
  MoveL 1605 to (0, -20.24, 3.4) mm, rotated rx 0 ry 0 rz 180 deg; joints [18.068, -54.765, 108.423, -157.951, 55.71, 77.147]
  MoveL 1606 to (-200, -20.24, 3.4) mm, rotated rx 0 ry 0 rz 180 deg; joints [20.902, -63.796, 124.368, -156.323, 62.677, 78.62]
  MoveL 1607 to (-200, -19.64, 3.4) mm, rotated rx 0 ry 0 rz 180 deg; joints [20.902, -63.762, 124.374, -156.332, 62.715, 78.639]
  MoveL 1608 to (0, -19.64, 3.4) mm, rotated rx 0 ry 0 rz 180 deg; joints [18.068, -54.737, 108.429, -157.96, 55.742, 77.162]
  MoveL 1609 to (0, -19.04, 3.4) mm, rotated rx 0 ry 0 rz 180 deg; joints [18.068, -54.708, 108.435, -157.969, 55.773, 77.178]
  MoveL 1610 to (-200, -19.04, 3.4) mm, rotated rx 0 ry 0 rz 180 deg; joints [20.902, -63.727, 124.38, -156.34, 62.752, 78.657]
  MoveL 1611 to (-200, -18.44, 3.4) mm, rotated rx 0 ry 0 rz 180 deg; joints [20.902, -63.693, 124.387, -156.348, 62.789, 78.675]
  MoveL 1612 to (0, -18.44, 3.4) mm, rotated rx 0 ry 0 rz 180 deg; joints [18.068, -54.68, 108.441, -157.978, 55.805, 77.193]
  MoveL 1613 to (0, -17.84, 3.4) mm, rotated rx 0 ry 0 rz 180 deg; joints [18.068, -54.652, 108.446, -157.986, 55.837, 77.208]
  MoveL 1614 to (-200, -17.84, 3.4) mm, rotated rx 0 ry 0 rz 180 deg; joints [20.902, -63.659, 124.393, -156.357, 62.826, 78.694]
  MoveL 1615 to (-200, -17.24, 3.4) mm, rotated rx 0 ry 0 rz 180 deg; joints [20.902, -63.624, 124.399, -156.365, 62.863, 78.712]
  MoveL 1616 to (0, -17.24, 3.4) mm, rotated rx 0 ry 0 rz 180 deg; joints [18.068, -54.623, 108.452, -157.995, 55.868, 77.224]
  MoveL 1617 to (0, -16.64, 3.4) mm, rotated rx 0 ry 0 rz 180 deg; joints [18.068, -54.595, 108.458, -158.004, 55.9, 77.239]
  MoveL 1618 to (-200, -16.64, 3.4) mm, rotated rx 0 ry 0 rz 180 deg; joints [20.902, -63.59, 124.405, -156.373, 62.901, 78.73]
  MoveL 1619 to (-200, -16.04, 3.4) mm, rotated rx 0 ry 0 rz 180 deg; joints [20.902, -63.555, 124.411, -156.382, 62.938, 78.749]
  MoveL 1620 to (0, -16.04, 3.4) mm, rotated rx 0 ry 0 rz 180 deg; joints [18.068, -54.567, 108.463, -158.012, 55.931, 77.255]
  MoveL 1621 to (0, -15.44, 3.4) mm, rotated rx 0 ry 0 rz 180 deg; joints [18.068, -54.539, 108.469, -158.021, 55.963, 77.27]
  MoveL 1622 to (-200, -15.44, 3.4) mm, rotated rx 0 ry 0 rz 180 deg; joints [20.902, -63.521, 124.418, -156.39, 62.975, 78.767]
  MoveL 1623 to (-200, -14.84, 3.4) mm, rotated rx 0 ry 0 rz 180 deg; joints [20.902, -63.487, 124.424, -156.398, 63.012, 78.785]
  MoveL 1624 to (0, -14.84, 3.4) mm, rotated rx 0 ry 0 rz 180 deg; joints [18.068, -54.51, 108.475, -158.029, 55.994, 77.285]
  MoveL 1625 to (0, -14.24, 3.4) mm, rotated rx 0 ry 0 rz 180 deg; joints [18.068, -54.482, 108.48, -158.038, 56.026, 77.301]
  MoveL 1626 to (-200, -14.24, 3.4) mm, rotated rx 0 ry 0 rz 180 deg; joints [20.902, -63.452, 124.43, -156.407, 63.049, 78.803]
  MoveL 1627 to (-200, -13.64, 3.4) mm, rotated rx 0 ry 0 rz 180 deg; joints [20.902, -63.418, 124.436, -156.415, 63.086, 78.821]
  MoveL 1628 to (0, -13.64, 3.4) mm, rotated rx 0 ry 0 rz 180 deg; joints [18.068, -54.453, 108.486, -158.046, 56.057, 77.316]
  MoveL 1629 to (0, -13.04, 3.4) mm, rotated rx 0 ry 0 rz 180 deg; joints [18.068, -54.425, 108.491, -158.055, 56.089, 77.331]
  MoveL 1630 to (-200, -13.04, 3.4) mm, rotated rx 0 ry 0 rz 180 deg; joints [20.902, -63.383, 124.442, -156.423, 63.124, 78.84]
  MoveL 1631 to (-200, -12.44, 3.4) mm, rotated rx 0 ry 0 rz 180 deg; joints [20.902, -63.349, 124.448, -156.431, 63.161, 78.858]
  MoveL 1632 to (0, -12.44, 3.4) mm, rotated rx 0 ry 0 rz 180 deg; joints [18.068, -54.397, 108.497, -158.063, 56.12, 77.347]
  MoveL 1633 to (0, -11.84, 3.4) mm, rotated rx 0 ry 0 rz 180 deg; joints [18.068, -54.368, 108.502, -158.072, 56.152, 77.362]
  MoveL 1634 to (-200, -11.84, 3.4) mm, rotated rx 0 ry 0 rz 180 deg; joints [20.902, -63.314, 124.454, -156.439, 63.198, 78.876]
  MoveL 1635 to (-200, -11.24, 3.4) mm, rotated rx 0 ry 0 rz 180 deg; joints [20.902, -63.279, 124.46, -156.448, 63.235, 78.894]
  MoveL 1636 to (0, -11.24, 3.4) mm, rotated rx 0 ry 0 rz 180 deg; joints [18.068, -54.34, 108.508, -158.08, 56.183, 77.377]
  MoveL 1637 to (0, -10.64, 3.4) mm, rotated rx 0 ry 0 rz 180 deg; joints [18.068, -54.311, 108.513, -158.089, 56.215, 77.392]
  MoveL 1638 to (-200, -10.64, 3.4) mm, rotated rx 0 ry 0 rz 180 deg; joints [20.902, -63.245, 124.466, -156.456, 63.272, 78.912]
  MoveL 1639 to (-200, -10.04, 3.4) mm, rotated rx 0 ry 0 rz 180 deg; joints [20.902, -63.21, 124.471, -156.464, 63.309, 78.93]
  MoveL 1640 to (0, -10.04, 3.4) mm, rotated rx 0 ry 0 rz 180 deg; joints [18.068, -54.283, 108.519, -158.097, 56.246, 77.407]
  MoveL 1641 to (0, -9.44, 3.4) mm, rotated rx 0 ry 0 rz 180 deg; joints [18.068, -54.254, 108.524, -158.106, 56.278, 77.423]
  MoveL 1642 to (-200, -9.44, 3.4) mm, rotated rx 0 ry 0 rz 180 deg; joints [20.902, -63.176, 124.477, -156.472, 63.346, 78.948]
  MoveL 1643 to (-200, -8.84, 3.4) mm, rotated rx 0 ry 0 rz 180 deg; joints [20.902, -63.141, 124.483, -156.48, 63.384, 78.966]
  MoveL 1644 to (0, -8.84, 3.4) mm, rotated rx 0 ry 0 rz 180 deg; joints [18.068, -54.226, 108.529, -158.114, 56.309, 77.438]
  MoveL 1645 to (0, -8.24, 3.4) mm, rotated rx 0 ry 0 rz 180 deg; joints [18.068, -54.197, 108.535, -158.123, 56.34, 77.453]
  MoveL 1646 to (-200, -8.24, 3.4) mm, rotated rx 0 ry 0 rz 180 deg; joints [20.902, -63.106, 124.489, -156.488, 63.421, 78.985]
  MoveL 1647 to (-200, -7.64, 3.4) mm, rotated rx 0 ry 0 rz 180 deg; joints [20.902, -63.071, 124.495, -156.496, 63.458, 79.003]
  MoveL 1648 to (0, -7.64, 3.4) mm, rotated rx 0 ry 0 rz 180 deg; joints [18.068, -54.168, 108.54, -158.131, 56.372, 77.468]
  MoveL 1649 to (0, -7.04, 3.4) mm, rotated rx 0 ry 0 rz 180 deg; joints [18.068, -54.14, 108.545, -158.139, 56.403, 77.483]
  MoveL 1650 to (-200, -7.04, 3.4) mm, rotated rx 0 ry 0 rz 180 deg; joints [20.902, -63.037, 124.5, -156.504, 63.495, 79.021]
  MoveL 1651 to (-200, -6.44, 3.4) mm, rotated rx 0 ry 0 rz 180 deg; joints [20.902, -63.002, 124.506, -156.512, 63.532, 79.039]
  MoveL 1652 to (0, -6.44, 3.4) mm, rotated rx 0 ry 0 rz 180 deg; joints [18.068, -54.111, 108.55, -158.148, 56.435, 77.498]
  MoveL 1653 to (0, -5.84, 3.4) mm, rotated rx 0 ry 0 rz 180 deg; joints [18.068, -54.083, 108.556, -158.156, 56.466, 77.514]
  MoveL 1654 to (-200, -5.84, 3.4) mm, rotated rx 0 ry 0 rz 180 deg; joints [20.902, -62.967, 124.512, -156.52, 63.569, 79.057]
  MoveL 1655 to (-200, -5.24, 3.4) mm, rotated rx 0 ry 0 rz 180 deg; joints [20.902, -62.932, 124.517, -156.528, 63.606, 79.075]
  MoveL 1656 to (0, -5.24, 3.4) mm, rotated rx 0 ry 0 rz 180 deg; joints [18.068, -54.054, 108.561, -158.164, 56.497, 77.529]
  MoveL 1657 to (0, -4.64, 3.4) mm, rotated rx 0 ry 0 rz 180 deg; joints [18.068, -54.025, 108.566, -158.173, 56.529, 77.544]
  MoveL 1658 to (-200, -4.64, 3.4) mm, rotated rx 0 ry 0 rz 180 deg; joints [20.902, -62.898, 124.523, -156.536, 63.643, 79.092]
  MoveL 1659 to (-200, -4.04, 3.4) mm, rotated rx 0 ry 0 rz 180 deg; joints [20.902, -62.863, 124.528, -156.544, 63.68, 79.11]
  MoveL 1660 to (0, -4.04, 3.4) mm, rotated rx 0 ry 0 rz 180 deg; joints [18.068, -53.997, 108.571, -158.181, 56.56, 77.559]
  MoveL 1661 to (0, -3.44, 3.4) mm, rotated rx 0 ry 0 rz 180 deg; joints [18.068, -53.968, 108.576, -158.189, 56.591, 77.574]
  MoveL 1662 to (-200, -3.44, 3.4) mm, rotated rx 0 ry 0 rz 180 deg; joints [20.902, -62.828, 124.534, -156.552, 63.717, 79.128]
  MoveL 1663 to (-200, -2.84, 3.4) mm, rotated rx 0 ry 0 rz 180 deg; joints [20.902, -62.793, 124.539, -156.56, 63.754, 79.146]
  MoveL 1664 to (0, -2.84, 3.4) mm, rotated rx 0 ry 0 rz 180 deg; joints [18.068, -53.939, 108.581, -158.198, 56.623, 77.589]
  MoveL 1665 to (0, -2.24, 3.4) mm, rotated rx 0 ry 0 rz 180 deg; joints [18.068, -53.91, 108.586, -158.206, 56.654, 77.604]
  MoveL 1666 to (-200, -2.24, 3.4) mm, rotated rx 0 ry 0 rz 180 deg; joints [20.902, -62.758, 124.545, -156.568, 63.791, 79.164]
  MoveL 1667 to (-200, -1.64, 3.4) mm, rotated rx 0 ry 0 rz 180 deg; joints [20.902, -62.723, 124.55, -156.576, 63.828, 79.182]
  MoveL 1668 to (0, -1.64, 3.4) mm, rotated rx 0 ry 0 rz 180 deg; joints [18.068, -53.882, 108.591, -158.214, 56.685, 77.619]
  MoveL 1669 to (0, -1.04, 3.4) mm, rotated rx 0 ry 0 rz 180 deg; joints [18.068, -53.853, 108.596, -158.222, 56.717, 77.634]
  MoveL 1670 to (-200, -1.04, 3.4) mm, rotated rx 0 ry 0 rz 180 deg; joints [20.902, -62.688, 124.555, -156.584, 63.865, 79.2]
  MoveL 1671 to (-200, -0.44, 3.4) mm, rotated rx 0 ry 0 rz 180 deg; joints [20.902, -62.653, 124.561, -156.592, 63.902, 79.218]
  MoveL 1672 to (0, -0.44, 3.4) mm, rotated rx 0 ry 0 rz 180 deg; joints [18.068, -53.824, 108.601, -158.231, 56.748, 77.649]
  MoveL 1673 to (0, 0, 3.4) mm, rotated rx 0 ry 0 rz 180 deg; joints [18.068, -53.803, 108.605, -158.237, 56.771, 77.66]
  MoveL 1674 to (-200, 0, 3.4) mm, rotated rx 0 ry 0 rz 180 deg; joints [20.902, -62.627, 124.565, -156.597, 63.929, 79.231]
  MoveL 1675 to (-200, 0, 3) mm, rotated rx 0 ry 0 rz 180 deg; joints [20.919, -62.621, 124.553, -156.578, 63.928, 79.22]
  MoveL 1676 to (0, 0, 3) mm, rotated rx 0 ry 0 rz 180 deg; joints [18.083, -53.797, 108.593, -158.218, 56.77, 77.648]
  MoveL 1677 to (0, -0.6, 3) mm, rotated rx 0 ry 0 rz 180 deg; joints [18.083, -53.826, 108.589, -158.21, 56.738, 77.633]
  MoveL 1678 to (-200, -0.6, 3) mm, rotated rx 0 ry 0 rz 180 deg; joints [20.919, -62.656, 124.548, -156.57, 63.891, 79.203]
  MoveL 1679 to (-200, -1.2, 3) mm, rotated rx 0 ry 0 rz 180 deg; joints [20.919, -62.691, 124.543, -156.562, 63.854, 79.185]
  MoveL 1680 to (0, -1.2, 3) mm, rotated rx 0 ry 0 rz 180 deg; joints [18.083, -53.855, 108.584, -158.201, 56.707, 77.618]
  MoveL 1681 to (0, -1.8, 3) mm, rotated rx 0 ry 0 rz 180 deg; joints [18.083, -53.883, 108.579, -158.193, 56.676, 77.603]
  MoveL 1682 to (-200, -1.8, 3) mm, rotated rx 0 ry 0 rz 180 deg; joints [20.919, -62.726, 124.537, -156.554, 63.817, 79.167]
  MoveL 1683 to (-200, -2.4, 3) mm, rotated rx 0 ry 0 rz 180 deg; joints [20.919, -62.761, 124.532, -156.546, 63.78, 79.149]
  MoveL 1684 to (0, -2.4, 3) mm, rotated rx 0 ry 0 rz 180 deg; joints [18.083, -53.912, 108.574, -158.185, 56.644, 77.588]
  MoveL 1685 to (0, -3, 3) mm, rotated rx 0 ry 0 rz 180 deg; joints [18.083, -53.941, 108.569, -158.177, 56.613, 77.573]
  MoveL 1686 to (-200, -3, 3) mm, rotated rx 0 ry 0 rz 180 deg; joints [20.919, -62.796, 124.526, -156.538, 63.743, 79.131]
  MoveL 1687 to (-200, -3.6, 3) mm, rotated rx 0 ry 0 rz 180 deg; joints [20.919, -62.83, 124.521, -156.53, 63.706, 79.113]
  MoveL 1688 to (0, -3.6, 3) mm, rotated rx 0 ry 0 rz 180 deg; joints [18.083, -53.969, 108.564, -158.168, 56.582, 77.558]
  MoveL 1689 to (0, -4.2, 3) mm, rotated rx 0 ry 0 rz 180 deg; joints [18.083, -53.998, 108.559, -158.16, 56.55, 77.543]
  MoveL 1690 to (-200, -4.2, 3) mm, rotated rx 0 ry 0 rz 180 deg; joints [20.919, -62.865, 124.515, -156.523, 63.669, 79.095]
  MoveL 1691 to (-200, -4.8, 3) mm, rotated rx 0 ry 0 rz 180 deg; joints [20.919, -62.9, 124.51, -156.515, 63.632, 79.077]
  MoveL 1692 to (0, -4.8, 3) mm, rotated rx 0 ry 0 rz 180 deg; joints [18.083, -54.027, 108.553, -158.152, 56.519, 77.528]
  MoveL 1693 to (0, -5.4, 3) mm, rotated rx 0 ry 0 rz 180 deg; joints [18.083, -54.055, 108.548, -158.143, 56.488, 77.513]
  MoveL 1694 to (-200, -5.4, 3) mm, rotated rx 0 ry 0 rz 180 deg; joints [20.919, -62.935, 124.504, -156.507, 63.595, 79.059]
  MoveL 1695 to (-200, -6, 3) mm, rotated rx 0 ry 0 rz 180 deg; joints [20.919, -62.97, 124.499, -156.499, 63.558, 79.041]
  MoveL 1696 to (0, -6, 3) mm, rotated rx 0 ry 0 rz 180 deg; joints [18.083, -54.084, 108.543, -158.135, 56.456, 77.497]
  MoveL 1697 to (0, -6.6, 3) mm, rotated rx 0 ry 0 rz 180 deg; joints [18.083, -54.113, 108.538, -158.127, 56.425, 77.482]
  MoveL 1698 to (-200, -6.6, 3) mm, rotated rx 0 ry 0 rz 180 deg; joints [20.919, -63.005, 124.493, -156.491, 63.521, 79.023]
  MoveL 1699 to (-200, -7.2, 3) mm, rotated rx 0 ry 0 rz 180 deg; joints [20.919, -63.039, 124.487, -156.482, 63.484, 79.005]
  MoveL 1700 to (0, -7.2, 3) mm, rotated rx 0 ry 0 rz 180 deg; joints [18.083, -54.141, 108.533, -158.118, 56.394, 77.467]
  MoveL 1701 to (0, -7.8, 3) mm, rotated rx 0 ry 0 rz 180 deg; joints [18.083, -54.17, 108.527, -158.11, 56.362, 77.452]
  MoveL 1702 to (-200, -7.8, 3) mm, rotated rx 0 ry 0 rz 180 deg; joints [20.919, -63.074, 124.482, -156.474, 63.447, 78.987]
  MoveL 1703 to (-200, -8.4, 3) mm, rotated rx 0 ry 0 rz 180 deg; joints [20.919, -63.109, 124.476, -156.466, 63.41, 78.969]
  MoveL 1704 to (0, -8.4, 3) mm, rotated rx 0 ry 0 rz 180 deg; joints [18.083, -54.198, 108.522, -158.102, 56.331, 77.437]
  MoveL 1705 to (0, -9, 3) mm, rotated rx 0 ry 0 rz 180 deg; joints [18.083, -54.227, 108.517, -158.093, 56.299, 77.422]
  MoveL 1706 to (-200, -9, 3) mm, rotated rx 0 ry 0 rz 180 deg; joints [20.919, -63.143, 124.47, -156.458, 63.373, 78.951]
  MoveL 1707 to (-200, -9.6, 3) mm, rotated rx 0 ry 0 rz 180 deg; joints [20.919, -63.178, 124.464, -156.45, 63.335, 78.933]
  MoveL 1708 to (0, -9.6, 3) mm, rotated rx 0 ry 0 rz 180 deg; joints [18.083, -54.256, 108.512, -158.085, 56.268, 77.407]
  MoveL 1709 to (0, -10.2, 3) mm, rotated rx 0 ry 0 rz 180 deg; joints [18.083, -54.284, 108.506, -158.076, 56.236, 77.391]
  MoveL 1710 to (-200, -10.2, 3) mm, rotated rx 0 ry 0 rz 180 deg; joints [20.919, -63.213, 124.458, -156.442, 63.298, 78.915]
  MoveL 1711 to (-200, -10.8, 3) mm, rotated rx 0 ry 0 rz 180 deg; joints [20.919, -63.247, 124.453, -156.434, 63.261, 78.897]
  MoveL 1712 to (0, -10.8, 3) mm, rotated rx 0 ry 0 rz 180 deg; joints [18.083, -54.313, 108.501, -158.068, 56.205, 77.376]
  MoveL 1713 to (0, -11.4, 3) mm, rotated rx 0 ry 0 rz 180 deg; joints [18.083, -54.341, 108.495, -158.059, 56.174, 77.361]
  MoveL 1714 to (-200, -11.4, 3) mm, rotated rx 0 ry 0 rz 180 deg; joints [20.919, -63.282, 124.447, -156.426, 63.224, 78.879]
  MoveL 1715 to (-200, -12, 3) mm, rotated rx 0 ry 0 rz 180 deg; joints [20.919, -63.316, 124.441, -156.418, 63.187, 78.861]
  MoveL 1716 to (0, -12, 3) mm, rotated rx 0 ry 0 rz 180 deg; joints [18.083, -54.37, 108.49, -158.051, 56.142, 77.346]
  MoveL 1717 to (0, -12.6, 3) mm, rotated rx 0 ry 0 rz 180 deg; joints [18.083, -54.398, 108.484, -158.042, 56.111, 77.33]
  MoveL 1718 to (-200, -12.6, 3) mm, rotated rx 0 ry 0 rz 180 deg; joints [20.919, -63.351, 124.435, -156.409, 63.15, 78.842]
  MoveL 1719 to (-200, -13.2, 3) mm, rotated rx 0 ry 0 rz 180 deg; joints [20.919, -63.386, 124.429, -156.401, 63.113, 78.824]
  MoveL 1720 to (0, -13.2, 3) mm, rotated rx 0 ry 0 rz 180 deg; joints [18.083, -54.426, 108.479, -158.034, 56.079, 77.315]
  MoveL 1721 to (0, -13.8, 3) mm, rotated rx 0 ry 0 rz 180 deg; joints [18.083, -54.455, 108.473, -158.025, 56.048, 77.3]
  MoveL 1722 to (-200, -13.8, 3) mm, rotated rx 0 ry 0 rz 180 deg; joints [20.919, -63.42, 124.423, -156.393, 63.076, 78.806]
  MoveL 1723 to (-200, -14.4, 3) mm, rotated rx 0 ry 0 rz 180 deg; joints [20.919, -63.455, 124.417, -156.385, 63.038, 78.788]
  MoveL 1724 to (0, -14.4, 3) mm, rotated rx 0 ry 0 rz 180 deg; joints [18.083, -54.483, 108.468, -158.017, 56.016, 77.284]
  MoveL 1725 to (0, -15, 3) mm, rotated rx 0 ry 0 rz 180 deg; joints [18.083, -54.512, 108.462, -158.008, 55.985, 77.269]
  MoveL 1726 to (-200, -15, 3) mm, rotated rx 0 ry 0 rz 180 deg; joints [20.919, -63.489, 124.411, -156.376, 63.001, 78.77]
  MoveL 1727 to (-200, -15.6, 3) mm, rotated rx 0 ry 0 rz 180 deg; joints [20.919, -63.523, 124.404, -156.368, 62.964, 78.751]
  MoveL 1728 to (0, -15.6, 3) mm, rotated rx 0 ry 0 rz 180 deg; joints [18.083, -54.54, 108.457, -157.999, 55.953, 77.254]
  MoveL 1729 to (0, -16.2, 3) mm, rotated rx 0 ry 0 rz 180 deg; joints [18.083, -54.568, 108.451, -157.991, 55.922, 77.238]
  MoveL 1730 to (-200, -16.2, 3) mm, rotated rx 0 ry 0 rz 180 deg; joints [20.919, -63.558, 124.398, -156.36, 62.927, 78.733]
  MoveL 1731 to (-200, -16.8, 3) mm, rotated rx 0 ry 0 rz 180 deg; joints [20.919, -63.592, 124.392, -156.351, 62.89, 78.715]
  MoveL 1732 to (0, -16.8, 3) mm, rotated rx 0 ry 0 rz 180 deg; joints [18.083, -54.597, 108.445, -157.982, 55.89, 77.223]
  MoveL 1733 to (0, -17.4, 3) mm, rotated rx 0 ry 0 rz 180 deg; joints [18.083, -54.625, 108.439, -157.974, 55.859, 77.208]
  MoveL 1734 to (-200, -17.4, 3) mm, rotated rx 0 ry 0 rz 180 deg; joints [20.919, -63.627, 124.386, -156.343, 62.853, 78.696]
  MoveL 1735 to (-200, -18, 3) mm, rotated rx 0 ry 0 rz 180 deg; joints [20.919, -63.661, 124.38, -156.335, 62.815, 78.678]
  MoveL 1736 to (0, -18, 3) mm, rotated rx 0 ry 0 rz 180 deg; joints [18.083, -54.653, 108.434, -157.965, 55.827, 77.192]
  MoveL 1737 to (0, -18.6, 3) mm, rotated rx 0 ry 0 rz 180 deg; joints [18.083, -54.681, 108.428, -157.956, 55.795, 77.177]
  MoveL 1738 to (-200, -18.6, 3) mm, rotated rx 0 ry 0 rz 180 deg; joints [20.919, -63.695, 124.373, -156.326, 62.778, 78.66]
  MoveL 1739 to (-200, -19.2, 3) mm, rotated rx 0 ry 0 rz 180 deg; joints [20.919, -63.73, 124.367, -156.318, 62.741, 78.641]
  MoveL 1740 to (0, -19.2, 3) mm, rotated rx 0 ry 0 rz 180 deg; joints [18.083, -54.71, 108.422, -157.948, 55.764, 77.161]
  MoveL 1741 to (0, -19.8, 3) mm, rotated rx 0 ry 0 rz 180 deg; joints [18.083, -54.738, 108.416, -157.939, 55.732, 77.146]
  MoveL 1742 to (-200, -19.8, 3) mm, rotated rx 0 ry 0 rz 180 deg; joints [20.919, -63.764, 124.361, -156.31, 62.704, 78.623]
  MoveL 1743 to (-200, -20.4, 3) mm, rotated rx 0 ry 0 rz 180 deg; joints [20.919, -63.798, 124.354, -156.301, 62.667, 78.605]
  MoveL 1744 to (0, -20.4, 3) mm, rotated rx 0 ry 0 rz 180 deg; joints [18.083, -54.766, 108.41, -157.93, 55.701, 77.13]
  MoveL 1745 to (0, -21, 3) mm, rotated rx 0 ry 0 rz 180 deg; joints [18.083, -54.794, 108.405, -157.921, 55.669, 77.115]
  MoveL 1746 to (-200, -21, 3) mm, rotated rx 0 ry 0 rz 180 deg; joints [20.919, -63.832, 124.348, -156.293, 62.629, 78.586]
  MoveL 1747 to (-200, -21.6, 3) mm, rotated rx 0 ry 0 rz 180 deg; joints [20.919, -63.867, 124.342, -156.284, 62.592, 78.568]
  MoveL 1748 to (0, -21.6, 3) mm, rotated rx 0 ry 0 rz 180 deg; joints [18.083, -54.822, 108.399, -157.913, 55.638, 77.099]
  MoveL 1749 to (0, -22.2, 3) mm, rotated rx 0 ry 0 rz 180 deg; joints [18.083, -54.851, 108.393, -157.904, 55.606, 77.084]
  MoveL 1750 to (-200, -22.2, 3) mm, rotated rx 0 ry 0 rz 180 deg; joints [20.919, -63.901, 124.335, -156.276, 62.555, 78.549]
  MoveL 1751 to (-200, -22.8, 3) mm, rotated rx 0 ry 0 rz 180 deg; joints [20.919, -63.935, 124.329, -156.267, 62.518, 78.531]
  MoveL 1752 to (0, -22.8, 3) mm, rotated rx 0 ry 0 rz 180 deg; joints [18.083, -54.879, 108.387, -157.895, 55.574, 77.068]
  MoveL 1753 to (0, -23.4, 3) mm, rotated rx 0 ry 0 rz 180 deg; joints [18.083, -54.907, 108.381, -157.886, 55.543, 77.052]
  MoveL 1754 to (-200, -23.4, 3) mm, rotated rx 0 ry 0 rz 180 deg; joints [20.919, -63.969, 124.322, -156.259, 62.48, 78.513]
  MoveL 1755 to (-200, -24, 3) mm, rotated rx 0 ry 0 rz 180 deg; joints [20.919, -64.003, 124.315, -156.25, 62.443, 78.494]
  MoveL 1756 to (0, -24, 3) mm, rotated rx 0 ry 0 rz 180 deg; joints [18.083, -54.935, 108.375, -157.877, 55.511, 77.037]
  MoveL 1757 to (0, -24.6, 3) mm, rotated rx 0 ry 0 rz 180 deg; joints [18.083, -54.963, 108.369, -157.869, 55.479, 77.021]
  MoveL 1758 to (-200, -24.6, 3) mm, rotated rx 0 ry 0 rz 180 deg; joints [20.919, -64.038, 124.309, -156.242, 62.406, 78.476]
  MoveL 1759 to (-200, -25.2, 3) mm, rotated rx 0 ry 0 rz 180 deg; joints [20.919, -64.072, 124.302, -156.233, 62.369, 78.457]
  MoveL 1760 to (0, -25.2, 3) mm, rotated rx 0 ry 0 rz 180 deg; joints [18.083, -54.991, 108.362, -157.86, 55.448, 77.006]
  MoveL 1761 to (0, -25.8, 3) mm, rotated rx 0 ry 0 rz 180 deg; joints [18.083, -55.019, 108.356, -157.851, 55.416, 76.99]
  MoveL 1762 to (-200, -25.8, 3) mm, rotated rx 0 ry 0 rz 180 deg; joints [20.919, -64.106, 124.296, -156.224, 62.331, 78.438]
  MoveL 1763 to (-200, -26.4, 3) mm, rotated rx 0 ry 0 rz 180 deg; joints [20.919, -64.14, 124.289, -156.216, 62.294, 78.42]
  MoveL 1764 to (0, -26.4, 3) mm, rotated rx 0 ry 0 rz 180 deg; joints [18.083, -55.047, 108.35, -157.842, 55.384, 76.974]
  MoveL 1765 to (0, -27, 3) mm, rotated rx 0 ry 0 rz 180 deg; joints [18.083, -55.075, 108.344, -157.833, 55.353, 76.959]
  MoveL 1766 to (-200, -27, 3) mm, rotated rx 0 ry 0 rz 180 deg; joints [20.919, -64.174, 124.282, -156.207, 62.257, 78.401]
  MoveL 1767 to (-200, -27.6, 3) mm, rotated rx 0 ry 0 rz 180 deg; joints [20.919, -64.208, 124.275, -156.198, 62.219, 78.383]
  MoveL 1768 to (0, -27.6, 3) mm, rotated rx 0 ry 0 rz 180 deg; joints [18.083, -55.103, 108.338, -157.824, 55.321, 76.943]
  MoveL 1769 to (0, -28.2, 3) mm, rotated rx 0 ry 0 rz 180 deg; joints [18.083, -55.131, 108.331, -157.815, 55.289, 76.927]
  MoveL 1770 to (-200, -28.2, 3) mm, rotated rx 0 ry 0 rz 180 deg; joints [20.919, -64.242, 124.269, -156.19, 62.182, 78.364]
  MoveL 1771 to (-200, -28.8, 3) mm, rotated rx 0 ry 0 rz 180 deg; joints [20.919, -64.276, 124.262, -156.181, 62.145, 78.346]
  MoveL 1772 to (0, -28.8, 3) mm, rotated rx 0 ry 0 rz 180 deg; joints [18.083, -55.159, 108.325, -157.806, 55.258, 76.912]
  MoveL 1773 to (0, -29.4, 3) mm, rotated rx 0 ry 0 rz 180 deg; joints [18.083, -55.187, 108.319, -157.797, 55.226, 76.896]
  MoveL 1774 to (-200, -29.4, 3) mm, rotated rx 0 ry 0 rz 180 deg; joints [20.919, -64.31, 124.255, -156.172, 62.107, 78.327]
  MoveL 1775 to (-200, -30, 3) mm, rotated rx 0 ry 0 rz 180 deg; joints [20.919, -64.344, 124.248, -156.164, 62.07, 78.308]
  MoveL 1776 to (0, -30, 3) mm, rotated rx 0 ry 0 rz 180 deg; joints [18.083, -55.215, 108.313, -157.788, 55.194, 76.88]
  MoveL 1777 to (0, -30.6, 3.02) mm, rotated rx 2.86 ry 0 rz 180 deg; joints [17.984, -56.104, 108.176, -157.631, 54.222, 79.337]
  MoveL 1778 to (-200, -30.6, 3.02) mm, rotated rx 2.86 ry 0 rz 180 deg; joints [20.807, -65.42, 124.096, -156.018, 60.924, 80.666]
  MoveL 1779 to (-200, -31.2, 3.06) mm, rotated rx 5.73 ry 0 rz 180 deg; joints [20.656, -66.484, 123.943, -155.906, 59.78, 83.045]
  MoveL 1780 to (0, -31.2, 3.06) mm, rotated rx 5.73 ry 0 rz 180 deg; joints [17.85, -56.984, 108.039, -157.507, 53.25, 81.815]
  MoveL 1781 to (0, -31.79, 3.13) mm, rotated rx 8.59 ry 0 rz 180 deg; joints [17.682, -57.853, 107.901, -157.419, 52.279, 84.319]
  MoveL 1782 to (-200, -31.79, 3.13) mm, rotated rx 8.59 ry 0 rz 180 deg; joints [20.466, -67.533, 123.787, -155.828, 58.637, 85.446]
  MoveL 1783 to (-200, -32.38, 3.24) mm, rotated rx 11.46 ry 0 rz 180 deg; joints [20.236, -68.567, 123.631, -155.788, 57.499, 87.876]
  MoveL 1784 to (0, -32.38, 3.24) mm, rotated rx 11.46 ry 0 rz 180 deg; joints [17.479, -58.71, 107.764, -157.368, 51.311, 86.852]
  MoveL 1785 to (0, -32.97, 3.37) mm, rotated rx 14.32 ry 0 rz 180 deg; joints [17.242, -59.552, 107.627, -157.357, 50.347, 89.418]
  MoveL 1786 to (-200, -32.97, 3.37) mm, rotated rx 14.32 ry 0 rz 180 deg; joints [19.967, -69.582, 123.474, -155.786, 56.366, 90.337]
  MoveL 1787 to (-200, -33.55, 3.54) mm, rotated rx 17.19 ry 0 rz 180 deg; joints [19.66, -70.577, 123.318, -155.826, 55.241, 92.834]
  MoveL 1788 to (0, -33.55, 3.54) mm, rotated rx 17.19 ry 0 rz 180 deg; joints [16.971, -60.377, 107.491, -157.387, 49.39, 92.02]
  MoveL 1789 to (0, -34.12, 3.73) mm, rotated rx 20.05 ry 0 rz 180 deg; joints [16.667, -61.185, 107.358, -157.462, 48.441, 94.662]
  MoveL 1790 to (-200, -34.12, 3.73) mm, rotated rx 20.05 ry 0 rz 180 deg; joints [19.315, -71.549, 123.163, -155.909, 54.126, 95.371]
  MoveL 1791 to (-200, -34.67, 3.95) mm, rotated rx 22.92 ry 0 rz 180 deg; joints [18.932, -72.497, 123.011, -156.039, 53.023, 97.952]
  MoveL 1792 to (0, -34.67, 3.95) mm, rotated rx 22.92 ry 0 rz 180 deg; joints [16.33, -61.973, 107.228, -157.583, 47.503, 97.346]
  MoveL 1793 to (0, -35.22, 4.2) mm, rotated rx 25.78 ry 0 rz 180 deg; joints [15.961, -62.74, 107.101, -157.753, 46.576, 100.078]
  MoveL 1794 to (-200, -35.22, 4.2) mm, rotated rx 25.78 ry 0 rz 180 deg; joints [18.511, -73.419, 122.861, -156.218, 51.934, 100.582]
  MoveL 1795 to (-200, -35.75, 4.47) mm, rotated rx 28.65 ry 0 rz 180 deg; joints [18.054, -74.313, 122.716, -156.449, 50.861, 103.265]
  MoveL 1796 to (0, -35.75, 4.47) mm, rotated rx 28.65 ry 0 rz 180 deg; joints [15.56, -63.484, 106.978, -157.974, 45.665, 102.861]
  MoveL 1797 to (0, -36.27, 4.77) mm, rotated rx 31.51 ry 0 rz 180 deg; joints [15.127, -64.203, 106.86, -158.251, 44.77, 105.699]
  MoveL 1798 to (-200, -36.27, 4.77) mm, rotated rx 31.51 ry 0 rz 180 deg; joints [17.561, -75.178, 122.575, -156.735, 49.807, 106.005]
  MoveL 1799 to (-200, -36.78, 5.1) mm, rotated rx 34.38 ry 0 rz 180 deg; joints [17.032, -76.011, 122.44, -157.08, 48.775, 108.807]
  MoveL 1800 to (0, -36.78, 5.1) mm, rotated rx 34.38 ry 0 rz 180 deg; joints [14.665, -64.897, 106.748, -158.584, 43.894, 108.595]
  MoveL 1801 to (0, -37.26, 5.45) mm, rotated rx 37.24 ry 0 rz 180 deg; joints [14.172, -65.564, 106.642, -158.978, 43.041, 111.553]
  MoveL 1802 to (-200, -37.26, 5.45) mm, rotated rx 37.24 ry 0 rz 180 deg; joints [16.469, -76.812, 122.312, -157.488, 47.766, 111.675]
  MoveL 1803 to (-200, -37.73, 5.82) mm, rotated rx 40.11 ry 0 rz 180 deg; joints [15.872, -77.578, 122.191, -157.96, 46.785, 114.613]
  MoveL 1804 to (0, -37.73, 5.82) mm, rotated rx 40.11 ry 0 rz 180 deg; joints [13.652, -66.203, 106.544, -159.434, 42.212, 114.577]
  MoveL 1805 to (0, -38.18, 6.22) mm, rotated rx 42.97 ry 0 rz 180 deg; joints [13.103, -66.811, 106.454, -159.956, 41.41, 117.669]
  MoveL 1806 to (-200, -38.18, 6.22) mm, rotated rx 42.97 ry 0 rz 180 deg; joints [15.242, -78.309, 122.079, -158.5, 45.835, 117.625]
  MoveL 1807 to (-200, -38.61, 6.64) mm, rotated rx 45.84 ry 0 rz 180 deg; joints [14.581, -79.002, 121.976, -159.112, 44.919, 120.715]
  MoveL 1808 to (0, -38.61, 6.64) mm, rotated rx 45.84 ry 0 rz 180 deg; joints [12.528, -67.389, 106.373, -160.545, 40.64, 120.832]
  MoveL 1809 to (0, -39.02, 7.08) mm, rotated rx 48.7 ry 0 rz 180 deg; joints [11.929, -67.935, 106.301, -161.204, 39.903, 124.068]
  MoveL 1810 to (-200, -39.02, 7.08) mm, rotated rx 48.7 ry 0 rz 180 deg; joints [13.891, -79.657, 121.883, -159.797, 44.041, 123.884]
  MoveL 1811 to (-200, -39.4, 7.54) mm, rotated rx 51.57 ry 0 rz 180 deg; joints [13.171, -80.272, 121.802, -160.559, 43.204, 127.138]
  MoveL 1812 to (0, -39.4, 7.54) mm, rotated rx 51.57 ry 0 rz 180 deg; joints [11.305, -68.448, 106.239, -161.933, 39.203, 127.379]
  MoveL 1813 to (0, -39.76, 8.02) mm, rotated rx 54.43 ry 0 rz 180 deg; joints [10.658, -68.926, 106.189, -162.733, 38.543, 130.767]
  MoveL 1814 to (-200, -39.76, 8.02) mm, rotated rx 54.43 ry 0 rz 180 deg; joints [12.425, -80.846, 121.732, -161.397, 42.413, 130.475]
  MoveL 1815 to (-200, -40.1, 8.52) mm, rotated rx 57.3 ry 0 rz 180 deg; joints [11.653, -81.378, 121.675, -162.314, 41.671, 133.899]
  MoveL 1816 to (0, -40.1, 8.52) mm, rotated rx 57.3 ry 0 rz 180 deg; joints [9.991, -69.369, 106.149, -163.605, 37.928, 134.23]
  MoveL 1817 to (0, -40.41, 9.03) mm, rotated rx 60.16 ry 0 rz 180 deg; joints [9.304, -69.775, 106.122, -164.548, 37.359, 137.769]
  MoveL 1818 to (-200, -40.41, 9.03) mm, rotated rx 60.16 ry 0 rz 180 deg; joints [10.857, -81.866, 121.632, -163.309, 40.983, 137.407]
  MoveL 1819 to (-200, -40.69, 9.56) mm, rotated rx 63.02 ry 0 rz 180 deg; joints [10.04, -82.31, 121.602, -164.381, 40.353, 140.998]
  MoveL 1820 to (0, -40.69, 9.56) mm, rotated rx 63.02 ry 0 rz 180 deg; joints [8.6, -70.145, 106.107, -165.558, 36.841, 141.379]
  MoveL 1821 to (0, -40.95, 10.1) mm, rotated rx 65.89 ry 0 rz 180 deg; joints [7.88, -70.476, 106.105, -166.635, 36.377, 145.061]
  MoveL 1822 to (-200, -40.95, 10.1) mm, rotated rx 65.89 ry 0 rz 180 deg; joints [9.203, -82.708, 121.588, -165.526, 39.785, 144.671]
  MoveL 1823 to (-200, -41.18, 10.65) mm, rotated rx 68.75 ry 0 rz 180 deg; joints [8.349, -83.06, 121.588, -166.742, 39.284, 148.42]
  MoveL 1824 to (0, -41.18, 10.65) mm, rotated rx 68.75 ry 0 rz 180 deg; joints [7.146, -70.769, 106.117, -167.773, 35.971, 148.808]
  MoveL 1825 to (0, -41.39, 11.22) mm, rotated rx 71.62 ry 0 rz 180 deg; joints [6.4, -71.022, 106.142, -168.968, 35.624, 152.615]
  MoveL 1826 to (-200, -41.39, 11.22) mm, rotated rx 71.62 ry 0 rz 180 deg; joints [7.48, -83.365, 121.604, -168.023, 38.853, 152.239]
  MoveL 1827 to (-200, -41.56, 11.79) mm, rotated rx 74.48 ry 0 rz 180 deg; joints [6.598, -83.622, 121.635, -169.362, 38.496, 156.122]
  MoveL 1828 to (0, -41.56, 11.79) mm, rotated rx 74.48 ry 0 rz 180 deg; joints [5.643, -71.235, 106.18, -170.212, 35.341, 156.475]
  MoveL 1829 to (0, -41.71, 12.37) mm, rotated rx 77.35 ry 0 rz 180 deg; joints [4.879, -71.408, 106.233, -171.498, 35.123, 160.378]
  MoveL 1830 to (-200, -41.71, 12.37) mm, rotated rx 77.35 ry 0 rz 180 deg; joints [5.707, -83.83, 121.683, -170.75, 38.217, 160.057]
  MoveL 1831 to (-200, -41.83, 12.96) mm, rotated rx 80.21 ry 0 rz 180 deg; joints [4.808, -83.989, 121.746, -172.179, 38.017, 164.038]
  MoveL 1832 to (0, -41.83, 12.96) mm, rotated rx 80.21 ry 0 rz 180 deg; joints [4.11, -71.539, 106.299, -172.818, 34.972, 164.318]
  MoveL 1833 to (0, -41.91, 13.55) mm, rotated rx 83.08 ry 0 rz 180 deg; joints [3.336, -71.629, 106.38, -174.161, 34.89, 168.284]
  MoveL 1834 to (-200, -41.91, 13.55) mm, rotated rx 83.08 ry 0 rz 180 deg; joints [3.904, -84.098, 121.826, -173.637, 37.899, 168.05]
  MoveL 1835 to (-200, -41.97, 14.15) mm, rotated rx 85.94 ry 0 rz 180 deg; joints [2.997, -84.157, 121.922, -175.113, 37.866, 172.082]
  MoveL 1836 to (0, -41.97, 14.15) mm, rotated rx 85.94 ry 0 rz 180 deg; joints [2.561, -71.677, 106.474, -175.518, 34.879, 172.265]
  MoveL 1837 to (0, -42, 14.75) mm, rotated rx 88.81 ry 0 rz 180 deg; joints [1.787, -71.683, 106.581, -176.878, 34.938, 176.248]
  MoveL 1838 to (-200, -42, 14.75) mm, rotated rx 88.81 ry 0 rz 180 deg; joints [2.092, -84.166, 122.033, -176.594, 37.917, 176.12]
  MoveL 1839 to (-200, -42, 15.35) mm, rotated rx 90 ry 0 rz 180 deg; joints [1.699, -84.155, 122.085, -177.237, 37.962, 177.821]
  MoveL 1840 to (0, -42, 15.35) mm, rotated rx 90 ry 0 rz 180 deg; joints [1.451, -71.674, 106.631, -177.468, 34.983, 177.925]
  MoveL 1841 to (0, -42, 15.95) mm, rotated rx 90 ry 0 rz 180 deg; joints [1.426, -71.675, 106.632, -177.512, 34.983, 177.961]
  MoveL 1842 to (-200, -42, 15.95) mm, rotated rx 90 ry 0 rz 180 deg; joints [1.67, -84.156, 122.086, -177.285, 37.961, 177.859]
  MoveL 1843 to (-200, -42, 16.55) mm, rotated rx 90 ry 0 rz 180 deg; joints [1.64, -84.157, 122.088, -177.333, 37.96, 177.896]
  MoveL 1844 to (0, -42, 16.55) mm, rotated rx 90 ry 0 rz 180 deg; joints [1.401, -71.676, 106.633, -177.555, 34.982, 177.996]
  MoveL 1845 to (0, -42, 17.15) mm, rotated rx 90 ry 0 rz 180 deg; joints [1.376, -71.676, 106.634, -177.599, 34.982, 178.032]
  MoveL 1846 to (-200, -42, 17.15) mm, rotated rx 90 ry 0 rz 180 deg; joints [1.611, -84.159, 122.089, -177.38, 37.959, 177.934]
  MoveL 1847 to (-200, -42, 17.75) mm, rotated rx 90 ry 0 rz 180 deg; joints [1.582, -84.16, 122.09, -177.428, 37.959, 177.971]
  MoveL 1848 to (0, -42, 17.75) mm, rotated rx 90 ry 0 rz 180 deg; joints [1.351, -71.677, 106.636, -177.643, 34.981, 178.068]
  MoveL 1849 to (0, -42, 18.35) mm, rotated rx 90 ry 0 rz 180 deg; joints [1.326, -71.678, 106.637, -177.686, 34.981, 178.104]
  MoveL 1850 to (-200, -42, 18.35) mm, rotated rx 90 ry 0 rz 180 deg; joints [1.552, -84.161, 122.091, -177.475, 37.958, 178.009]
  MoveL 1851 to (-200, -42, 18.95) mm, rotated rx 90 ry 0 rz 180 deg; joints [1.523, -84.162, 122.092, -177.523, 37.957, 178.047]
  MoveL 1852 to (0, -42, 18.95) mm, rotated rx 90 ry 0 rz 180 deg; joints [1.301, -71.679, 106.638, -177.73, 34.98, 178.14]
  MoveL 1853 to (0, -42, 19.55) mm, rotated rx 90 ry 0 rz 180 deg; joints [1.276, -71.68, 106.639, -177.774, 34.98, 178.175]
  MoveL 1854 to (-200, -42, 19.55) mm, rotated rx 90 ry 0 rz 180 deg; joints [1.494, -84.163, 122.094, -177.571, 37.956, 178.084]
  MoveL 1855 to (-200, -42, 20.15) mm, rotated rx 90 ry 0 rz 180 deg; joints [1.465, -84.164, 122.095, -177.618, 37.955, 178.122]
  MoveL 1856 to (0, -42, 20.15) mm, rotated rx 90 ry 0 rz 180 deg; joints [1.251, -71.681, 106.64, -177.817, 34.979, 178.211]
  MoveL 1857 to (0, -42, 20.75) mm, rotated rx 90 ry 0 rz 180 deg; joints [1.226, -71.681, 106.641, -177.861, 34.979, 178.247]
  MoveL 1858 to (-200, -42, 20.75) mm, rotated rx 90 ry 0 rz 180 deg; joints [1.435, -84.165, 122.096, -177.666, 37.954, 178.159]
  MoveL 1859 to (-200, -42, 21.35) mm, rotated rx 90 ry 0 rz 180 deg; joints [1.406, -84.166, 122.097, -177.714, 37.953, 178.197]
  MoveL 1860 to (0, -42, 21.35) mm, rotated rx 90 ry 0 rz 180 deg; joints [1.201, -71.682, 106.642, -177.905, 34.978, 178.283]
  MoveL 1861 to (0, -42, 21.95) mm, rotated rx 90 ry 0 rz 180 deg; joints [1.176, -71.683, 106.643, -177.948, 34.978, 178.319]
  MoveL 1862 to (-200, -42, 21.95) mm, rotated rx 90 ry 0 rz 180 deg; joints [1.377, -84.167, 122.098, -177.761, 37.953, 178.234]
  MoveL 1863 to (-200, -42, 22.55) mm, rotated rx 90 ry 0 rz 180 deg; joints [1.347, -84.167, 122.099, -177.809, 37.952, 178.272]
  MoveL 1864 to (0, -42, 22.55) mm, rotated rx 90 ry 0 rz 180 deg; joints [1.151, -71.684, 106.644, -177.992, 34.977, 178.354]
  MoveL 1865 to (0, -42, 23.15) mm, rotated rx 90 ry 0 rz 180 deg; joints [1.126, -71.684, 106.645, -178.036, 34.977, 178.39]
  MoveL 1866 to (-200, -42, 23.15) mm, rotated rx 90 ry 0 rz 180 deg; joints [1.318, -84.168, 122.1, -177.857, 37.951, 178.31]
  MoveL 1867 to (-200, -42, 23.75) mm, rotated rx 90 ry 0 rz 180 deg; joints [1.289, -84.169, 122.101, -177.904, 37.95, 178.347]
  MoveL 1868 to (0, -42, 23.75) mm, rotated rx 90 ry 0 rz 180 deg; joints [1.101, -71.685, 106.646, -178.079, 34.976, 178.426]
  MoveL 1869 to (0, -42, 24.35) mm, rotated rx 90 ry 0 rz 180 deg; joints [1.076, -71.686, 106.647, -178.123, 34.976, 178.462]
  MoveL 1870 to (-200, -42, 24.35) mm, rotated rx 90 ry 0 rz 180 deg; joints [1.259, -84.17, 122.102, -177.952, 37.95, 178.385]
  MoveL 1871 to (-200, -42, 24.95) mm, rotated rx 90 ry 0 rz 180 deg; joints [1.23, -84.171, 122.103, -178, 37.949, 178.422]
  MoveL 1872 to (0, -42, 24.95) mm, rotated rx 90 ry 0 rz 180 deg; joints [1.051, -71.687, 106.648, -178.167, 34.975, 178.498]
  MoveL 1873 to (0, -42, 25.55) mm, rotated rx 90 ry 0 rz 180 deg; joints [1.026, -71.687, 106.649, -178.21, 34.975, 178.533]
  MoveL 1874 to (-200, -42, 25.55) mm, rotated rx 90 ry 0 rz 180 deg; joints [1.201, -84.172, 122.104, -178.047, 37.948, 178.46]
  MoveL 1875 to (-200, -42, 26.15) mm, rotated rx 90 ry 0 rz 180 deg; joints [1.171, -84.173, 122.105, -178.095, 37.947, 178.498]
  MoveL 1876 to (0, -42, 26.15) mm, rotated rx 90 ry 0 rz 180 deg; joints [1.001, -71.688, 106.65, -178.254, 34.975, 178.569]
  MoveL 1877 to (0, -42, 26.75) mm, rotated rx 90 ry 0 rz 180 deg; joints [0.976, -71.689, 106.651, -178.298, 34.974, 178.605]
  MoveL 1878 to (-200, -42, 26.75) mm, rotated rx 90 ry 0 rz 180 deg; joints [1.142, -84.173, 122.106, -178.143, 37.947, 178.535]
  MoveL 1879 to (-200, -42, 27.35) mm, rotated rx 90 ry 0 rz 180 deg; joints [1.113, -84.174, 122.106, -178.19, 37.946, 178.573]
  MoveL 1880 to (0, -42, 27.35) mm, rotated rx 90 ry 0 rz 180 deg; joints [0.951, -71.689, 106.652, -178.342, 34.974, 178.641]
  MoveL 1881 to (0, -42, 27.95) mm, rotated rx 90 ry 0 rz 180 deg; joints [0.925, -71.69, 106.653, -178.385, 34.973, 178.677]
  MoveL 1882 to (-200, -42, 27.95) mm, rotated rx 90 ry 0 rz 180 deg; joints [1.083, -84.175, 122.107, -178.238, 37.945, 178.61]
  MoveL 1883 to (-200, -42, 28.55) mm, rotated rx 90 ry 0 rz 180 deg; joints [1.054, -84.176, 122.108, -178.286, 37.945, 178.648]
  MoveL 1884 to (0, -42, 28.55) mm, rotated rx 90 ry 0 rz 180 deg; joints [0.9, -71.69, 106.653, -178.429, 34.973, 178.713]
  MoveL 1885 to (0, -42, 29.15) mm, rotated rx 90 ry 0 rz 180 deg; joints [0.875, -71.691, 106.654, -178.473, 34.973, 178.748]
  MoveL 1886 to (-200, -42, 29.15) mm, rotated rx 90 ry 0 rz 180 deg; joints [1.025, -84.176, 122.109, -178.333, 37.944, 178.685]
  MoveL 1887 to (-200, -42, 29.75) mm, rotated rx 90 ry 0 rz 180 deg; joints [0.995, -84.177, 122.11, -178.381, 37.944, 178.723]
  MoveL 1888 to (0, -42, 29.75) mm, rotated rx 90 ry 0 rz 180 deg; joints [0.85, -71.692, 106.655, -178.516, 34.972, 178.784]
  MoveL 1889 to (0, -42, 30.35) mm, rotated rx 90 ry 0 rz 180 deg; joints [0.825, -71.692, 106.656, -178.56, 34.972, 178.82]
  MoveL 1890 to (-200, -42, 30.35) mm, rotated rx 90 ry 0 rz 180 deg; joints [0.966, -84.178, 122.11, -178.429, 37.943, 178.761]
  MoveL 1891 to (-200, -42, 30.95) mm, rotated rx 90 ry 0 rz 180 deg; joints [0.937, -84.178, 122.111, -178.476, 37.943, 178.798]
  MoveL 1892 to (0, -42, 30.95) mm, rotated rx 90 ry 0 rz 180 deg; joints [0.8, -71.693, 106.656, -178.604, 34.972, 178.856]
  MoveL 1893 to (0, -42, 31.55) mm, rotated rx 90 ry 0 rz 180 deg; joints [0.775, -71.693, 106.657, -178.647, 34.971, 178.892]
  MoveL 1894 to (-200, -42, 31.55) mm, rotated rx 90 ry 0 rz 180 deg; joints [0.907, -84.179, 122.112, -178.524, 37.942, 178.836]
  MoveL 1895 to (-200, -42, 32.15) mm, rotated rx 90 ry 0 rz 180 deg; joints [0.878, -84.179, 122.112, -178.572, 37.941, 178.874]
  MoveL 1896 to (0, -42, 32.15) mm, rotated rx 90 ry 0 rz 180 deg; joints [0.75, -71.694, 106.658, -178.691, 34.971, 178.927]
  MoveL 1897 to (0, -42, 32.75) mm, rotated rx 90 ry 0 rz 180 deg; joints [0.725, -71.694, 106.658, -178.735, 34.971, 178.963]
  MoveL 1898 to (-200, -42, 32.75) mm, rotated rx 90 ry 0 rz 180 deg; joints [0.849, -84.18, 122.113, -178.619, 37.941, 178.911]
  MoveL 1899 to (-200, -42, 33.35) mm, rotated rx 90 ry 0 rz 180 deg; joints [0.819, -84.181, 122.114, -178.667, 37.941, 178.949]
  MoveL 1900 to (0, -42, 33.35) mm, rotated rx 90 ry 0 rz 180 deg; joints [0.7, -71.694, 106.659, -178.779, 34.971, 178.999]
  MoveL 1901 to (0, -42, 33.95) mm, rotated rx 90 ry 0 rz 180 deg; joints [0.675, -71.695, 106.66, -178.822, 34.97, 179.035]
  MoveL 1902 to (-200, -42, 33.95) mm, rotated rx 90 ry 0 rz 180 deg; joints [0.79, -84.181, 122.114, -178.715, 37.94, 178.986]
  MoveL 1903 to (-200, -42, 34.55) mm, rotated rx 90 ry 0 rz 180 deg; joints [0.761, -84.182, 122.115, -178.763, 37.94, 179.024]
  MoveL 1904 to (0, -42, 34.55) mm, rotated rx 90 ry 0 rz 180 deg; joints [0.65, -71.695, 106.66, -178.866, 34.97, 179.071]
  MoveL 1905 to (0, -42, 35.15) mm, rotated rx 90 ry 0 rz 180 deg; joints [0.625, -71.696, 106.661, -178.91, 34.97, 179.107]
  MoveL 1906 to (-200, -42, 35.15) mm, rotated rx 90 ry 0 rz 180 deg; joints [0.731, -84.182, 122.115, -178.81, 37.939, 179.062]
  MoveL 1907 to (-200, -42, 35.75) mm, rotated rx 90 ry 0 rz 180 deg; joints [0.702, -84.183, 122.116, -178.858, 37.939, 179.099]
  MoveL 1908 to (0, -42, 35.75) mm, rotated rx 90 ry 0 rz 180 deg; joints [0.6, -71.696, 106.661, -178.953, 34.97, 179.142]
  MoveL 1909 to (0, -42, 36.35) mm, rotated rx 90 ry 0 rz 180 deg; joints [0.575, -71.697, 106.662, -178.997, 34.969, 179.178]
  MoveL 1910 to (-200, -42, 36.35) mm, rotated rx 90 ry 0 rz 180 deg; joints [0.673, -84.183, 122.116, -178.906, 37.938, 179.137]
  MoveL 1911 to (-200, -42, 36.95) mm, rotated rx 90 ry 0 rz 180 deg; joints [0.643, -84.184, 122.117, -178.953, 37.938, 179.174]
  MoveL 1912 to (0, -42, 36.95) mm, rotated rx 90 ry 0 rz 180 deg; joints [0.55, -71.697, 106.662, -179.041, 34.969, 179.214]
  MoveL 1913 to (0, -42, 37.55) mm, rotated rx 90 ry 0 rz 180 deg; joints [0.525, -71.697, 106.663, -179.085, 34.969, 179.25]
  MoveL 1914 to (-200, -42, 37.55) mm, rotated rx 90 ry 0 rz 180 deg; joints [0.614, -84.184, 122.117, -179.001, 37.938, 179.212]
  MoveL 1915 to (-200, -42, 38.15) mm, rotated rx 90 ry 0 rz 180 deg; joints [0.585, -84.184, 122.118, -179.049, 37.937, 179.25]
  MoveL 1916 to (0, -42, 38.15) mm, rotated rx 90 ry 0 rz 180 deg; joints [0.5, -71.698, 106.663, -179.128, 34.969, 179.286]
  MoveL 1917 to (0, -42, 38.75) mm, rotated rx 90 ry 0 rz 180 deg; joints [0.475, -71.698, 106.664, -179.172, 34.968, 179.321]
  MoveL 1918 to (-200, -42, 38.75) mm, rotated rx 90 ry 0 rz 180 deg; joints [0.556, -84.185, 122.118, -179.096, 37.937, 179.287]
  MoveL 1919 to (-200, -42, 39.35) mm, rotated rx 90 ry 0 rz 180 deg; joints [0.526, -84.185, 122.119, -179.144, 37.937, 179.325]
  MoveL 1920 to (0, -42, 39.35) mm, rotated rx 90 ry 0 rz 180 deg; joints [0.449, -71.698, 106.664, -179.216, 34.968, 179.357]
  MoveL 1921 to (0, -42, 39.95) mm, rotated rx 90 ry 0 rz 180 deg; joints [0.424, -71.698, 106.664, -179.259, 34.968, 179.393]
  MoveL 1922 to (-200, -42, 39.95) mm, rotated rx 90 ry 0 rz 180 deg; joints [0.497, -84.185, 122.119, -179.192, 37.936, 179.363]
  MoveL 1923 to (-200, -42, 40.55) mm, rotated rx 90 ry 0 rz 180 deg; joints [0.468, -84.186, 122.119, -179.24, 37.936, 179.4]
  MoveL 1924 to (0, -42, 40.55) mm, rotated rx 90 ry 0 rz 180 deg; joints [0.399, -71.699, 106.665, -179.303, 34.968, 179.429]
  MoveL 1925 to (0, -42, 41.15) mm, rotated rx 90 ry 0 rz 180 deg; joints [0.374, -71.699, 106.665, -179.347, 34.968, 179.465]
  MoveL 1926 to (-200, -42, 41.15) mm, rotated rx 90 ry 0 rz 180 deg; joints [0.438, -84.186, 122.12, -179.287, 37.936, 179.438]
  MoveL 1927 to (-200, -42, 41.75) mm, rotated rx 90 ry 0 rz 180 deg; joints [0.409, -84.186, 122.12, -179.335, 37.936, 179.475]
  MoveL 1928 to (0, -42, 41.75) mm, rotated rx 90 ry 0 rz 180 deg; joints [0.349, -71.699, 106.665, -179.391, 34.968, 179.501]
  MoveL 1929 to (0, -42, 42.35) mm, rotated rx 90 ry 0 rz 180 deg; joints [0.324, -71.699, 106.666, -179.434, 34.967, 179.536]
  MoveL 1930 to (-200, -42, 42.35) mm, rotated rx 90 ry 0 rz 180 deg; joints [0.38, -84.187, 122.12, -179.383, 37.935, 179.513]
  MoveL 1931 to (-200, -42, 42.95) mm, rotated rx 90 ry 0 rz 180 deg; joints [0.35, -84.187, 122.121, -179.43, 37.935, 179.551]
  MoveL 1932 to (0, -42, 42.95) mm, rotated rx 90 ry 0 rz 180 deg; joints [0.299, -71.7, 106.666, -179.478, 34.967, 179.572]
  MoveL 1933 to (0, -42, 43.55) mm, rotated rx 90 ry 0 rz 180 deg; joints [0.274, -71.7, 106.666, -179.522, 34.967, 179.608]
  MoveL 1934 to (-200, -42, 43.55) mm, rotated rx 90 ry 0 rz 180 deg; joints [0.321, -84.187, 122.121, -179.478, 37.935, 179.588]
  MoveL 1935 to (-200, -42, 44.15) mm, rotated rx 90 ry 0 rz 180 deg; joints [0.292, -84.187, 122.121, -179.526, 37.935, 179.626]
  MoveL 1936 to (0, -42, 44.15) mm, rotated rx 90 ry 0 rz 180 deg; joints [0.249, -71.7, 106.666, -179.565, 34.967, 179.644]
  MoveL 1937 to (0, -42, 44.75) mm, rotated rx 90 ry 0 rz 180 deg; joints [0.224, -71.7, 106.667, -179.609, 34.967, 179.68]
  MoveL 1938 to (-200, -42, 44.75) mm, rotated rx 90 ry 0 rz 180 deg; joints [0.262, -84.188, 122.121, -179.574, 37.935, 179.664]
  MoveL 1939 to (-200, -41.99, 45.35) mm, rotated rx 91.67 ry 0 rz 180 deg; joints [-0.277, -84.139, 122.178, 179.551, 38.039, -177.973]
  MoveL 1940 to (0, -41.99, 45.35) mm, rotated rx 91.67 ry 0 rz 180 deg; joints [-0.236, -71.659, 106.719, 179.588, 35.06, -177.99]
  MoveL 1941 to (0, -41.96, 45.95) mm, rotated rx 94.54 ry 0 rz 180 deg; joints [-1.002, -71.556, 106.819, 178.265, 35.275, -174.045]
  MoveL 1942 to (-200, -41.96, 45.95) mm, rotated rx 94.54 ry 0 rz 180 deg; joints [-1.173, -84.016, 122.286, 178.106, 38.286, -173.975]
  MoveL 1943 to (-200, -41.9, 46.55) mm, rotated rx 97.4 ry 0 rz 180 deg; joints [-2.06, -83.842, 122.409, 176.698, 38.614, -170.016]
  MoveL 1944 to (0, -41.9, 46.55) mm, rotated rx 97.4 ry 0 rz 180 deg; joints [-1.76, -71.411, 106.932, 176.973, 35.559, -170.133]
  MoveL 1945 to (0, -41.81, 47.14) mm, rotated rx 100.27 ry 0 rz 180 deg; joints [-2.508, -71.224, 107.057, 175.722, 35.909, -166.264]
  MoveL 1946 to (-200, -41.81, 47.14) mm, rotated rx 100.27 ry 0 rz 180 deg; joints [-2.935, -83.618, 122.547, 175.335, 39.022, -166.105]
  MoveL 1947 to (-200, -41.69, 47.73) mm, rotated rx 103.13 ry 0 rz 180 deg; joints [-3.795, -83.343, 122.698, 174.028, 39.507, -162.254]
  MoveL 1948 to (0, -41.69, 47.73) mm, rotated rx 103.13 ry 0 rz 180 deg; joints [-3.243, -70.995, 107.193, 174.519, 36.323, -162.447]
  MoveL 1949 to (0, -41.53, 48.31) mm, rotated rx 106 ry 0 rz 180 deg; joints [-3.965, -70.725, 107.34, 173.372, 36.798, -158.687]
  MoveL 1950 to (-200, -41.53, 48.31) mm, rotated rx 106 ry 0 rz 180 deg; joints [-4.639, -83.019, 122.861, 172.782, 40.067, -158.467]
  MoveL 1951 to (-200, -41.36, 48.88) mm, rotated rx 108.86 ry 0 rz 180 deg; joints [-5.463, -82.646, 123.037, 171.605, 40.696, -154.754]
  MoveL 1952 to (0, -41.36, 48.88) mm, rotated rx 108.86 ry 0 rz 180 deg; joints [-4.67, -70.415, 107.497, 172.284, 37.333, -154.99]
  MoveL 1953 to (0, -41.15, 49.44) mm, rotated rx 111.73 ry 0 rz 180 deg; joints [-5.357, -70.064, 107.663, 171.262, 37.923, -151.36]
  MoveL 1954 to (-200, -41.15, 49.44) mm, rotated rx 111.73 ry 0 rz 180 deg; joints [-6.265, -82.223, 123.224, 170.501, 41.392, -151.118]
  MoveL 1955 to (-200, -40.91, 49.99) mm, rotated rx 114.59 ry 0 rz 180 deg; joints [-7.044, -81.753, 123.421, 169.472, 42.151, -147.563]
  MoveL 1956 to (0, -40.91, 49.99) mm, rotated rx 114.59 ry 0 rz 180 deg; joints [-6.025, -69.674, 107.838, 170.307, 38.565, -147.801]
  MoveL 1957 to (0, -40.65, 50.53) mm, rotated rx 117.46 ry 0 rz 180 deg; joints [-6.671, -69.244, 108.02, 169.422, 39.256, -144.316]
  MoveL 1958 to (-200, -40.65, 50.53) mm, rotated rx 117.46 ry 0 rz 180 deg; joints [-7.796, -81.236, 123.626, 168.52, 42.968, -144.091]
  MoveL 1959 to (-200, -40.36, 51.06) mm, rotated rx 120.32 ry 0 rz 180 deg; joints [-8.521, -80.672, 123.84, 167.647, 43.838, -140.702]
  MoveL 1960 to (0, -40.36, 51.06) mm, rotated rx 120.32 ry 0 rz 180 deg; joints [-7.294, -68.777, 108.209, 168.607, 39.992, -140.903]
  MoveL 1961 to (0, -40.04, 51.57) mm, rotated rx 123.19 ry 0 rz 180 deg; joints [-7.892, -68.272, 108.403, 167.863, 40.77, -137.563]
  MoveL 1962 to (-200, -40.04, 51.57) mm, rotated rx 123.19 ry 0 rz 180 deg; joints [-9.217, -80.062, 124.06, 166.851, 44.759, -137.396]
  MoveL 1963 to (-200, -39.7, 52.06) mm, rotated rx 126.05 ry 0 rz 180 deg; joints [-9.882, -79.408, 124.286, 166.132, 45.725, -134.17]
  MoveL 1964 to (0, -39.7, 52.06) mm, rotated rx 126.05 ry 0 rz 180 deg; joints [-8.464, -67.731, 108.602, 167.188, 41.587, -134.296]
  MoveL 1965 to (0, -39.34, 52.54) mm, rotated rx 128.92 ry 0 rz 180 deg; joints [-9.009, -67.154, 108.804, 166.582, 42.438, -131.099]
  MoveL 1966 to (-200, -39.34, 52.54) mm, rotated rx 128.92 ry 0 rz 180 deg; joints [-10.514, -78.711, 124.516, 165.487, 46.733, -131.023]
  MoveL 1967 to (-200, -38.95, 52.99) mm, rotated rx 131.78 ry 0 rz 180 deg; joints [-11.112, -77.972, 124.75, 164.915, 47.779, -127.953]
  MoveL 1968 to (0, -38.95, 52.99) mm, rotated rx 131.78 ry 0 rz 180 deg; joints [-9.525, -66.544, 109.009, 166.044, 43.321, -127.972]
  MoveL 1969 to (0, -38.54, 53.43) mm, rotated rx 134.65 ry 0 rz 180 deg; joints [-10.011, -65.9, 109.216, 165.57, 44.233, -124.909]
  MoveL 1970 to (-200, -38.54, 53.43) mm, rotated rx 134.65 ry 0 rz 180 deg; joints [-11.676, -77.192, 124.985, 164.412, 48.859, -124.954]
  MoveL 1971 to (-200, -38.11, 53.85) mm, rotated rx 137.51 ry 0 rz 180 deg; joints [-12.203, -76.373, 125.22, 163.975, 49.969, -122.023]
  MoveL 1972 to (0, -38.11, 53.85) mm, rotated rx 137.51 ry 0 rz 180 deg; joints [-10.467, -65.225, 109.423, 165.158, 45.17, -121.908]
  MoveL 1973 to (0, -37.65, 54.24) mm, rotated rx 140.38 ry 0 rz 180 deg; joints [-10.89, -64.519, 109.629, 164.807, 46.129, -118.966]
  MoveL 1974 to (-200, -37.65, 54.24) mm, rotated rx 140.38 ry 0 rz 180 deg; joints [-12.693, -75.516, 125.456, 163.602, 51.107, -119.157]
  MoveL 1975 to (-200, -37.18, 54.61) mm, rotated rx 143.24 ry 0 rz 180 deg; joints [-13.145, -74.624, 125.689, 163.289, 52.268, -116.35]
  MoveL 1976 to (0, -37.18, 54.61) mm, rotated rx 143.24 ry 0 rz 180 deg; joints [-11.282, -63.784, 109.834, 164.513, 47.107, -116.081]
  MoveL 1977 to (0, -36.69, 54.96) mm, rotated rx 146.1 ry 0 rz 180 deg; joints [-11.64, -63.022, 110.036, 164.273, 48.102, -113.246]
  MoveL 1978 to (-200, -36.69, 54.96) mm, rotated rx 146.1 ry 0 rz 180 deg; joints [-13.558, -73.697, 125.919, 163.033, 53.449, -113.598]
  MoveL 1979 to (-200, -36.19, 55.28) mm, rotated rx 148.97 ry 0 rz 180 deg; joints [-13.931, -72.737, 126.145, 162.832, 54.649, -110.896]
  MoveL 1980 to (0, -36.19, 55.28) mm, rotated rx 148.97 ry 0 rz 180 deg; joints [-11.964, -62.234, 110.234, 164.086, 49.111, -110.459]
  MoveL 1981 to (0, -35.66, 55.58) mm, rotated rx 151.83 ry 0 rz 180 deg; joints [-12.253, -61.422, 110.429, 163.948, 50.131, -107.715]
  MoveL 1982 to (-200, -35.66, 55.58) mm, rotated rx 151.83 ry 0 rz 180 deg; joints [-14.265, -71.747, 126.366, 162.681, 55.863, -108.24]
  MoveL 1983 to (-200, -35.13, 55.85) mm, rotated rx 154.7 ry 0 rz 180 deg; joints [-14.557, -70.729, 126.58, 162.578, 57.089, -105.625]
  MoveL 1984 to (0, -35.13, 55.85) mm, rotated rx 154.7 ry 0 rz 180 deg; joints [-12.507, -60.588, 110.618, 163.857, 51.16, -105.012]
  MoveL 1985 to (0, -34.58, 56.09) mm, rotated rx 157.56 ry 0 rz 180 deg; joints [-12.726, -59.733, 110.8, 163.81, 52.195, -102.346]
  MoveL 1986 to (-200, -34.58, 56.09) mm, rotated rx 157.56 ry 0 rz 180 deg; joints [-14.809, -69.686, 126.787, 162.522, 58.324, -103.048]
  MoveL 1987 to (-200, -34.02, 56.31) mm, rotated rx 160.43 ry 0 rz 180 deg; joints [-15.02, -68.618, 126.986, 162.509, 59.567, -100.503]
  MoveL 1988 to (0, -34.02, 56.31) mm, rotated rx 160.43 ry 0 rz 180 deg; joints [-12.909, -58.86, 110.976, 163.807, 53.235, -99.712]
  MoveL 1989 to (0, -33.45, 56.49) mm, rotated rx 163.29 ry 0 rz 180 deg; joints [-13.056, -57.97, 111.145, 163.844, 54.276, -97.106]
  MoveL 1990 to (-200, -33.45, 56.49) mm, rotated rx 163.29 ry 0 rz 180 deg; joints [-15.188, -67.528, 127.176, 162.537, 60.813, -97.985]
  MoveL 1991 to (-200, -32.87, 56.65) mm, rotated rx 166.16 ry 0 rz 180 deg; joints [-15.315, -66.42, 127.356, 162.604, 62.061, -95.491]
  MoveL 1992 to (0, -32.87, 56.65) mm, rotated rx 166.16 ry 0 rz 180 deg; joints [-13.166, -57.065, 111.305, 163.919, 55.317, -94.526]
  MoveL 1993 to (0, -32.28, 56.78) mm, rotated rx 169.02 ry 0 rz 180 deg; joints [-13.24, -56.148, 111.457, 164.031, 56.356, -91.968]
  MoveL 1994 to (-200, -32.28, 56.78) mm, rotated rx 169.02 ry 0 rz 180 deg; joints [-15.4, -65.296, 127.526, 162.709, 63.308, -93.017]
  MoveL 1995 to (-200, -31.69, 56.88) mm, rotated rx 171.89 ry 0 rz 180 deg; joints [-15.442, -64.158, 127.684, 162.85, 64.551, -90.559]
  MoveL 1996 to (0, -31.69, 56.88) mm, rotated rx 171.89 ry 0 rz 180 deg; joints [-13.277, -55.221, 111.599, 164.179, 57.39, -89.43]
  MoveL 1997 to (0, -31.1, 56.95) mm, rotated rx 174.75 ry 0 rz 180 deg; joints [-13.277, -54.287, 111.732, 164.36, 58.418, -86.907]
  MoveL 1998 to (-200, -31.1, 56.95) mm, rotated rx 174.75 ry 0 rz 180 deg; joints [-15.442, -63.01, 127.831, 163.026, 65.79, -88.113]
  MoveL 1999 to (-200, -30.5, 56.99) mm, rotated rx 177.62 ry 0 rz 180 deg; joints [-15.4, -61.853, 127.966, 163.235, 67.02, -85.675]
  MoveL 2000 to (0, -30.5, 56.99) mm, rotated rx 177.62 ry 0 rz 180 deg; joints [-13.241, -53.346, 111.854, 164.574, 59.437, -84.396]
  MoveL 2001 to (0, -29.9, 57) mm, rotated rx 180 ry 0 rz 180 deg; joints [-13.182, -52.556, 111.949, 164.777, 60.282, -82.317]
  MoveL 2002 to (-200, -29.9, 57) mm, rotated rx 180 ry 0 rz 180 deg; joints [-15.333, -60.881, 128.069, 163.435, 68.043, -83.654]
  MoveL 2003 to (-200, -29.3, 57) mm, rotated rx 180 ry 0 rz 180 deg; joints [-15.333, -60.842, 128.071, 163.439, 68.082, -83.666]
  MoveL 2004 to (0, -29.3, 57) mm, rotated rx 180 ry 0 rz 180 deg; joints [-13.182, -52.525, 111.951, 164.782, 60.314, -82.327]
  MoveL 2005 to (0, -28.7, 57) mm, rotated rx 180 ry 0 rz 180 deg; joints [-13.182, -52.493, 111.953, 164.787, 60.346, -82.337]
  MoveL 2006 to (-200, -28.7, 57) mm, rotated rx 180 ry 0 rz 180 deg; joints [-15.333, -60.804, 128.073, 163.444, 68.121, -83.679]
  MoveL 2007 to (-200, -28.1, 57) mm, rotated rx 180 ry 0 rz 180 deg; joints [-15.333, -60.765, 128.076, 163.449, 68.16, -83.691]
  MoveL 2008 to (0, -28.1, 57) mm, rotated rx 180 ry 0 rz 180 deg; joints [-13.182, -52.462, 111.955, 164.792, 60.379, -82.347]
  MoveL 2009 to (0, -27.5, 57) mm, rotated rx 180 ry 0 rz 180 deg; joints [-13.182, -52.43, 111.957, 164.797, 60.411, -82.357]
  MoveL 2010 to (-200, -27.5, 57) mm, rotated rx 180 ry 0 rz 180 deg; joints [-15.333, -60.727, 128.078, 163.453, 68.199, -83.704]
  MoveL 2011 to (-200, -26.9, 57) mm, rotated rx 180 ry 0 rz 180 deg; joints [-15.333, -60.688, 128.08, 163.458, 68.239, -83.716]
  MoveL 2012 to (0, -26.9, 57) mm, rotated rx 180 ry 0 rz 180 deg; joints [-13.182, -52.399, 111.959, 164.802, 60.443, -82.367]
  MoveL 2013 to (0, -26.3, 57) mm, rotated rx 180 ry 0 rz 180 deg; joints [-13.182, -52.368, 111.961, 164.807, 60.475, -82.377]
  MoveL 2014 to (-200, -26.3, 57) mm, rotated rx 180 ry 0 rz 180 deg; joints [-15.333, -60.65, 128.082, 163.463, 68.278, -83.729]
  MoveL 2015 to (-200, -25.7, 57) mm, rotated rx 180 ry 0 rz 180 deg; joints [-15.333, -60.611, 128.084, 163.467, 68.317, -83.741]
  MoveL 2016 to (0, -25.7, 57) mm, rotated rx 180 ry 0 rz 180 deg; joints [-13.182, -52.336, 111.963, 164.812, 60.508, -82.388]
  MoveL 2017 to (0, -25.1, 57) mm, rotated rx 180 ry 0 rz 180 deg; joints [-13.182, -52.305, 111.965, 164.816, 60.54, -82.398]
  MoveL 2018 to (-200, -25.1, 57) mm, rotated rx 180 ry 0 rz 180 deg; joints [-15.333, -60.572, 128.086, 163.472, 68.356, -83.754]
  MoveL 2019 to (-200, -24.5, 57) mm, rotated rx 180 ry 0 rz 180 deg; joints [-15.333, -60.534, 128.089, 163.476, 68.395, -83.766]
  MoveL 2020 to (0, -24.5, 57) mm, rotated rx 180 ry 0 rz 180 deg; joints [-13.182, -52.273, 111.967, 164.821, 60.572, -82.408]
  MoveL 2021 to (0, -23.9, 57) mm, rotated rx 180 ry 0 rz 180 deg; joints [-13.182, -52.242, 111.969, 164.826, 60.604, -82.418]
  MoveL 2022 to (-200, -23.9, 57) mm, rotated rx 180 ry 0 rz 180 deg; joints [-15.333, -60.495, 128.091, 163.481, 68.434, -83.779]
  MoveL 2023 to (-200, -23.3, 57) mm, rotated rx 180 ry 0 rz 180 deg; joints [-15.333, -60.456, 128.093, 163.486, 68.473, -83.791]
  MoveL 2024 to (0, -23.3, 57) mm, rotated rx 180 ry 0 rz 180 deg; joints [-13.182, -52.21, 111.97, 164.831, 60.637, -82.428]
  MoveL 2025 to (0, -22.7, 57) mm, rotated rx 180 ry 0 rz 180 deg; joints [-13.182, -52.179, 111.972, 164.836, 60.669, -82.438]
  MoveL 2026 to (-200, -22.7, 57) mm, rotated rx 180 ry 0 rz 180 deg; joints [-15.333, -60.418, 128.095, 163.49, 68.512, -83.803]
  MoveL 2027 to (-200, -22.1, 57) mm, rotated rx 180 ry 0 rz 180 deg; joints [-15.333, -60.379, 128.097, 163.495, 68.551, -83.816]
  MoveL 2028 to (0, -22.1, 57) mm, rotated rx 180 ry 0 rz 180 deg; joints [-13.182, -52.147, 111.974, 164.841, 60.701, -82.448]
  MoveL 2029 to (0, -21.5, 57) mm, rotated rx 180 ry 0 rz 180 deg; joints [-13.182, -52.115, 111.976, 164.846, 60.733, -82.458]
  MoveL 2030 to (-200, -21.5, 57) mm, rotated rx 180 ry 0 rz 180 deg; joints [-15.333, -60.34, 128.098, 163.499, 68.59, -83.828]
  MoveL 2031 to (-200, -20.9, 57) mm, rotated rx 180 ry 0 rz 180 deg; joints [-15.333, -60.301, 128.1, 163.504, 68.629, -83.841]
  MoveL 2032 to (0, -20.9, 57) mm, rotated rx 180 ry 0 rz 180 deg; joints [-13.182, -52.084, 111.977, 164.851, 60.765, -82.468]
  MoveL 2033 to (0, -20.3, 57) mm, rotated rx 180 ry 0 rz 180 deg; joints [-13.182, -52.052, 111.979, 164.856, 60.797, -82.478]
  MoveL 2034 to (-200, -20.3, 57) mm, rotated rx 180 ry 0 rz 180 deg; joints [-15.333, -60.263, 128.102, 163.508, 68.668, -83.853]
  MoveL 2035 to (-200, -19.7, 57) mm, rotated rx 180 ry 0 rz 180 deg; joints [-15.333, -60.224, 128.104, 163.513, 68.707, -83.865]
  MoveL 2036 to (0, -19.7, 57) mm, rotated rx 180 ry 0 rz 180 deg; joints [-13.182, -52.021, 111.981, 164.861, 60.829, -82.488]
  MoveL 2037 to (0, -19.1, 57) mm, rotated rx 180 ry 0 rz 180 deg; joints [-13.182, -51.989, 111.982, 164.865, 60.862, -82.497]
  MoveL 2038 to (-200, -19.1, 57) mm, rotated rx 180 ry 0 rz 180 deg; joints [-15.333, -60.185, 128.106, 163.517, 68.746, -83.878]
  MoveL 2039 to (-200, -18.5, 57) mm, rotated rx 180 ry 0 rz 180 deg; joints [-15.333, -60.146, 128.108, 163.522, 68.785, -83.89]
  MoveL 2040 to (0, -18.5, 57) mm, rotated rx 180 ry 0 rz 180 deg; joints [-13.182, -51.957, 111.984, 164.87, 60.894, -82.507]
  MoveL 2041 to (0, -17.9, 57) mm, rotated rx 180 ry 0 rz 180 deg; joints [-13.182, -51.926, 111.985, 164.875, 60.926, -82.517]
  MoveL 2042 to (-200, -17.9, 57) mm, rotated rx 180 ry 0 rz 180 deg; joints [-15.333, -60.107, 128.109, 163.526, 68.824, -83.902]
  MoveL 2043 to (-200, -17.3, 57) mm, rotated rx 180 ry 0 rz 180 deg; joints [-15.333, -60.068, 128.111, 163.531, 68.862, -83.915]
  MoveL 2044 to (0, -17.3, 57) mm, rotated rx 180 ry 0 rz 180 deg; joints [-13.182, -51.894, 111.987, 164.88, 60.958, -82.527]
  MoveL 2045 to (0, -16.7, 57) mm, rotated rx 180 ry 0 rz 180 deg; joints [-13.182, -51.862, 111.988, 164.885, 60.99, -82.537]
  MoveL 2046 to (-200, -16.7, 57) mm, rotated rx 180 ry 0 rz 180 deg; joints [-15.333, -60.03, 128.113, 163.535, 68.901, -83.927]
  MoveL 2047 to (-200, -16.1, 57) mm, rotated rx 180 ry 0 rz 180 deg; joints [-15.333, -59.991, 128.114, 163.539, 68.94, -83.939]
  MoveL 2048 to (0, -16.1, 57) mm, rotated rx 180 ry 0 rz 180 deg; joints [-13.182, -51.83, 111.99, 164.889, 61.022, -82.547]
  MoveL 2049 to (0, -15.5, 57) mm, rotated rx 180 ry 0 rz 180 deg; joints [-13.182, -51.799, 111.991, 164.894, 61.054, -82.557]
  MoveL 2050 to (-200, -15.5, 57) mm, rotated rx 180 ry 0 rz 180 deg; joints [-15.333, -59.952, 128.116, 163.544, 68.979, -83.952]
  MoveL 2051 to (-200, -14.9, 57) mm, rotated rx 180 ry 0 rz 180 deg; joints [-15.333, -59.913, 128.117, 163.548, 69.018, -83.964]
  MoveL 2052 to (0, -14.9, 57) mm, rotated rx 180 ry 0 rz 180 deg; joints [-13.182, -51.767, 111.993, 164.899, 61.086, -82.567]
  MoveL 2053 to (0, -14.3, 57) mm, rotated rx 180 ry 0 rz 180 deg; joints [-13.182, -51.735, 111.994, 164.904, 61.118, -82.577]
  MoveL 2054 to (-200, -14.3, 57) mm, rotated rx 180 ry 0 rz 180 deg; joints [-15.333, -59.874, 128.119, 163.553, 69.057, -83.976]
  MoveL 2055 to (-200, -13.7, 57) mm, rotated rx 180 ry 0 rz 180 deg; joints [-15.333, -59.835, 128.12, 163.557, 69.096, -83.989]
  MoveL 2056 to (0, -13.7, 57) mm, rotated rx 180 ry 0 rz 180 deg; joints [-13.182, -51.703, 111.995, 164.909, 61.15, -82.587]
  MoveL 2057 to (0, -13.1, 57) mm, rotated rx 180 ry 0 rz 180 deg; joints [-13.182, -51.672, 111.997, 164.913, 61.182, -82.596]
  MoveL 2058 to (-200, -13.1, 57) mm, rotated rx 180 ry 0 rz 180 deg; joints [-15.333, -59.796, 128.122, 163.561, 69.134, -84.001]
